(* Logix 5000 project; controller NWGG 1756-L72 rev 35.12; software revision 35.00; part 2 of 19 *)
(* tags used below, declared in another part *)
   T22 : TIMER[100];
   T4 : TIMER[100];

ADD_ON_INSTRUCTION Loadout_K_Valve_Control   (* revision 1.0 *)
VAR_IN_OUT
   K_Valve : udt_Loadout_K_Valve; {required}
   ALM_Clean_Pos_Failed : ALARM_DIGITAL; {required}
   ALM_Treat_Pos_Failed : ALARM_DIGITAL; {required}
   Treat_Position_Input : BOOL; {required}
   Clean_Position_Input : BOOL; {required}
   Clean_Gate_Relay : BOOL; {required}
   Treat_Gate_Relay : BOOL; {required}
END_VAR
VAR
   Clean_Pos_Failed_ACK : BOOL; {access None}
   Treat_Pos_Failedt_ACK : BOOL; {access None}
END_VAR

ROUTINE Logic   (* ladder *)
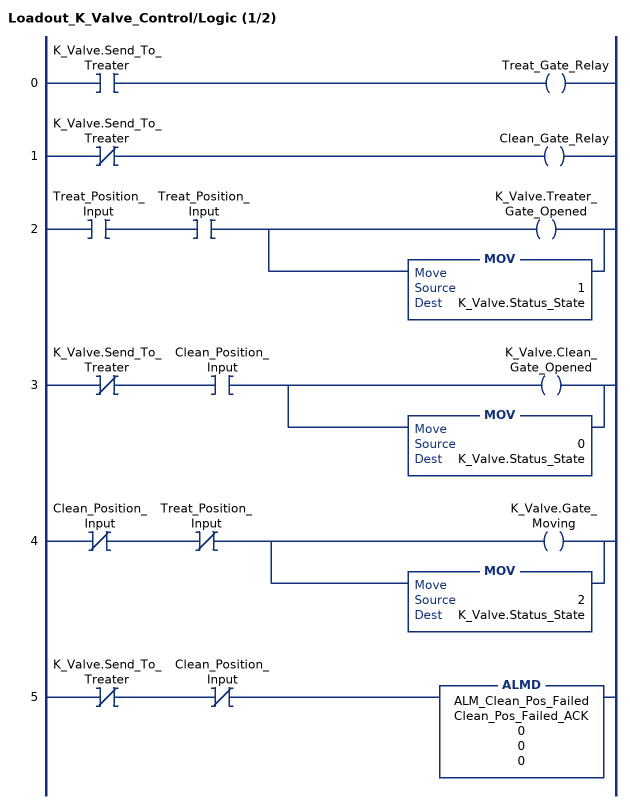
   0: XIC(K_Valve.Send_To_Treater)OTE(Treat_Gate_Relay);
   1: XIO(K_Valve.Send_To_Treater)OTE(Clean_Gate_Relay);
   2: XIC(Treat_Position_Input)XIC(Treat_Position_Input)[OTE(K_Valve.Treater_Gate_Opened) ,MOV(1,K_Valve.Status_State) ];
   3: XIO(K_Valve.Send_To_Treater)XIC(Clean_Position_Input)[OTE(K_Valve.Clean_Gate_Opened) ,MOV(0,K_Valve.Status_State) ];
   4: XIO(Clean_Position_Input)XIO(Treat_Position_Input)[OTE(K_Valve.Gate_Moving) ,MOV(2,K_Valve.Status_State) ];
   5: XIO(K_Valve.Send_To_Treater)XIO(Clean_Position_Input)ALMD(ALM_Clean_Pos_Failed,Clean_Pos_Failed_ACK,0,0,0);
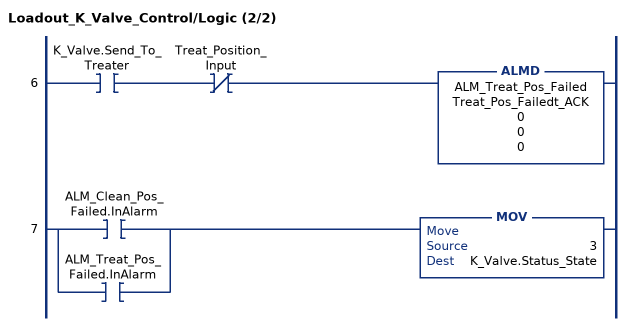
   6: XIC(K_Valve.Send_To_Treater)XIO(Treat_Position_Input)ALMD(ALM_Treat_Pos_Failed,Treat_Pos_Failedt_ACK,0,0,0);
   7: [XIC(ALM_Clean_Pos_Failed.InAlarm) ,XIC(ALM_Treat_Pos_Failed.InAlarm) ]MOV(3,K_Valve.Status_State);
END_ROUTINE
END_ADD_ON_INSTRUCTION

ADD_ON_INSTRUCTION Motor_Control   (* revision 1.0 *)
VAR_IN_OUT
   Motor_Contact : BOOL; {required}
END_VAR
VAR_INPUT
   Spd_20_Pct : BOOL; {required}
   Spd_10_Pct : BOOL; {required}
END_VAR
VAR_OUTPUT
   Running : BOOL; {access Read Only, required}
END_VAR
VAR_IN_OUT
   Motor_Alarm_SPD20 : ALARM_DIGITAL; {required}
   Motor_Alarm_SPD10 : ALARM_DIGITAL; {required}
   Motor_Alarm_Stopped_Over_Amps : ALARM_DIGITAL; {required}
   Motor_Start : udt_Motor_Start; {required}
END_VAR
VAR_INPUT
   Plugged_Sensor : BOOL; {required}
END_VAR
VAR_IN_OUT
   Motor_Alarm_Plugged : ALARM_DIGITAL; {required}
END_VAR
VAR_INPUT
   Motor_Amps : REAL; {required}
END_VAR
VAR_IN_OUT
   Motor_Config : udt_Motor_Config; {required}
   Motor_Starting : BOOL; {required}
   Motor_Alarm_Wont_Start : ALARM_DIGITAL; {required}
END_VAR
VAR_OUTPUT
   In_Alarm : BOOL; {access Read Only}
END_VAR
VAR_IN_OUT
   Treat_Batch_Status : DINT; {required}
   Clean_Batch_Status : DINT; {required}
   Transfer_Batch_Status : DINT; {required}
END_VAR
VAR_OUTPUT
   Motor_Batch_Ready : BOOL; {access Read Only}
END_VAR
VAR_IN_OUT
   Manual_Mode : BOOL; {required}
   InterLocked_Belt : BOOL; {required}
END_VAR
VAR_OUTPUT
   Motor_Batch_Ready_Clean : BOOL; {access Read Only}
   Motor_Batch_Ready_Treat : BOOL; {access Read Only}
   Motor_Batch_Ready_Transfer : BOOL; {access Read Only}
END_VAR
VAR
   TMR_BELT_SPD20 : TIMER := (PRE := 2000); {access None}
   TMR_AMP_INRUSH : TIMER := (PRE := 2000); {access None}
   Alm_Spd20_AK : BOOL; {access None}
   Alm_Spd10_AK : BOOL; {access None}
   Alm_Plugged_AK : BOOL; {access None}
   Alm_OVR_AMP_AK : BOOL; {access None}
   Stop_Motor_Plugged : BOOL; {access None}
   Stop_Motor_SLP20 : BOOL; {access None}
   Stop_Motor : BOOL; {access None}
   Stop_Motor_Ovr_Amp : BOOL; {access None}
   TMR_BELT_SPD10 : TIMER := (PRE := 2000); {access None}
   Alm_Wont_Start_AK : BOOL; {access None}
   Req_Motor_Start : BOOL; {access None}
   tmr_Auto_Stop_Delay : TIMER; {access None}
END_VAR

ROUTINE Logic   (* ladder *)
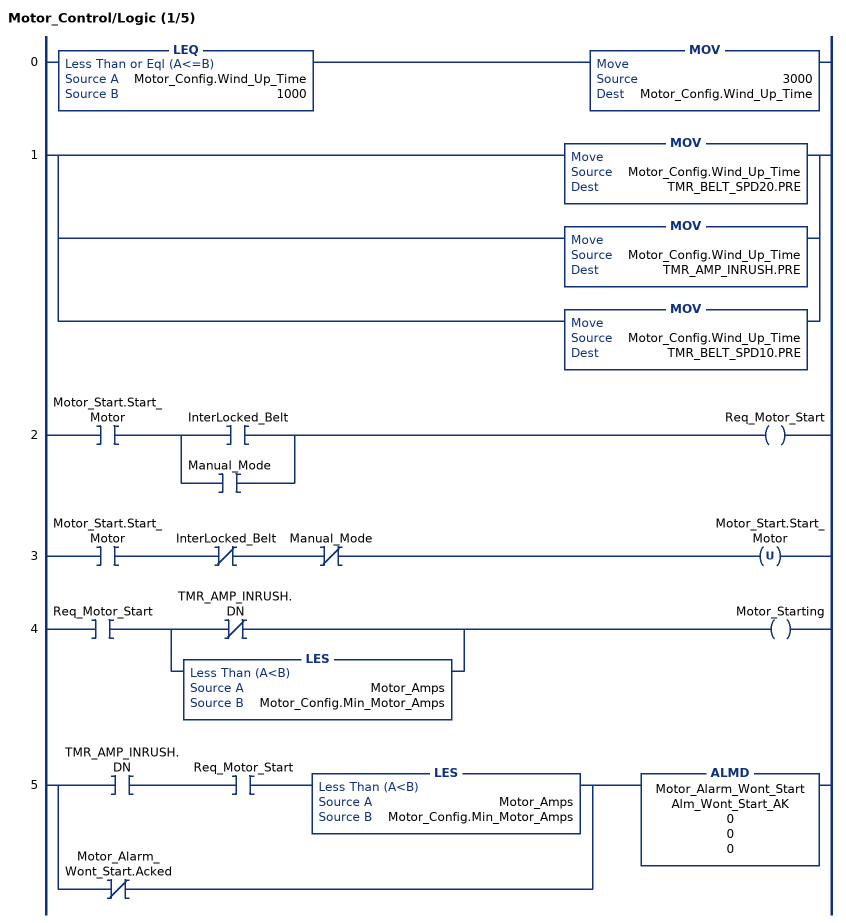
   0: LEQ(Motor_Config.Wind_Up_Time,1000)MOV(3000,Motor_Config.Wind_Up_Time);
   1: [MOV(Motor_Config.Wind_Up_Time,TMR_BELT_SPD20.PRE) ,MOV(Motor_Config.Wind_Up_Time,TMR_AMP_INRUSH.PRE) ,MOV(Motor_Config.Wind_Up_Time,TMR_BELT_SPD10.PRE) ];
   2: XIC(Motor_Start.Start_Motor)[XIC(InterLocked_Belt) ,XIC(Manual_Mode) ]OTE(Req_Motor_Start);
   3: XIC(Motor_Start.Start_Motor)XIO(InterLocked_Belt)XIO(Manual_Mode)OTU(Motor_Start.Start_Motor);
   4: XIC(Req_Motor_Start)[XIO(TMR_AMP_INRUSH.DN) ,LES(Motor_Amps,Motor_Config.Min_Motor_Amps) ]OTE(Motor_Starting);
   5: [XIC(TMR_AMP_INRUSH.DN) XIC(Req_Motor_Start) LES(Motor_Amps,Motor_Config.Min_Motor_Amps) ,XIO(Motor_Alarm_Wont_Start.Acked) ]ALMD(Motor_Alarm_Wont_Start,Alm_Wont_Start_AK,0,0,0);
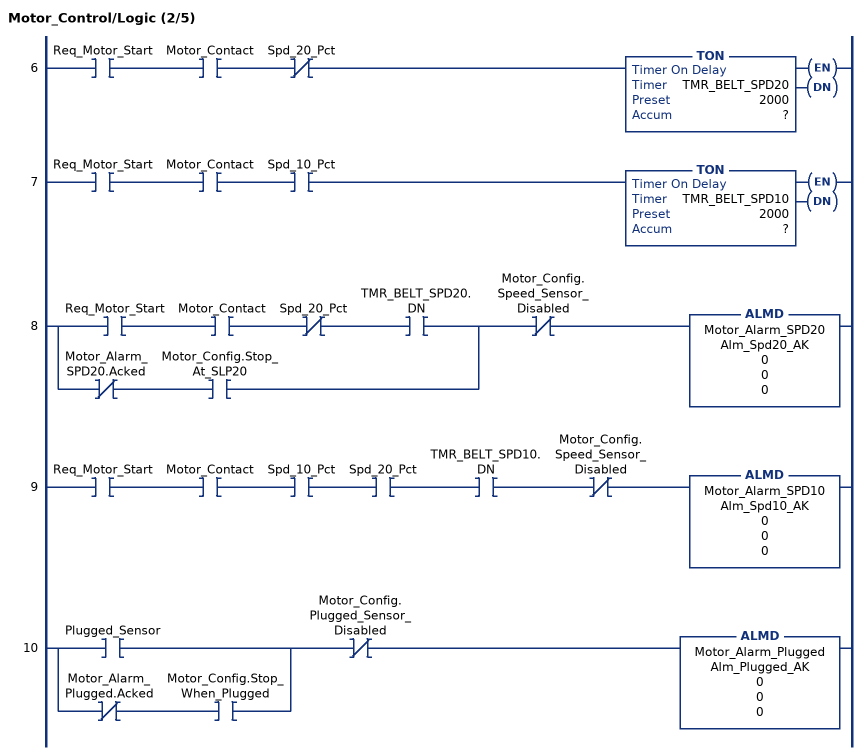
   6: XIC(Req_Motor_Start)XIC(Motor_Contact)XIO(Spd_20_Pct)TON(TMR_BELT_SPD20,?,?);
   7: XIC(Req_Motor_Start)XIC(Motor_Contact)XIC(Spd_10_Pct)TON(TMR_BELT_SPD10,?,?);
   8: [XIC(Req_Motor_Start) XIC(Motor_Contact) XIO(Spd_20_Pct) XIC(TMR_BELT_SPD20.DN) ,XIO(Motor_Alarm_SPD20.Acked) XIC(Motor_Config.Stop_At_SLP20) ]XIO(Motor_Config.Speed_Sensor_Disabled)ALMD(Motor_Alarm_SPD20,Alm_Spd20_AK,0,0,0);
   9: XIC(Req_Motor_Start)XIC(Motor_Contact)XIC(Spd_10_Pct)XIC(Spd_20_Pct)XIC(TMR_BELT_SPD10.DN)XIO(Motor_Config.Speed_Sensor_Disabled)ALMD(Motor_Alarm_SPD10,Alm_Spd10_AK,0,0,0);
   10: [XIC(Plugged_Sensor) ,XIO(Motor_Alarm_Plugged.Acked) XIC(Motor_Config.Stop_When_Plugged) ]XIO(Motor_Config.Plugged_Sensor_Disabled)ALMD(Motor_Alarm_Plugged,Alm_Plugged_AK,0,0,0);
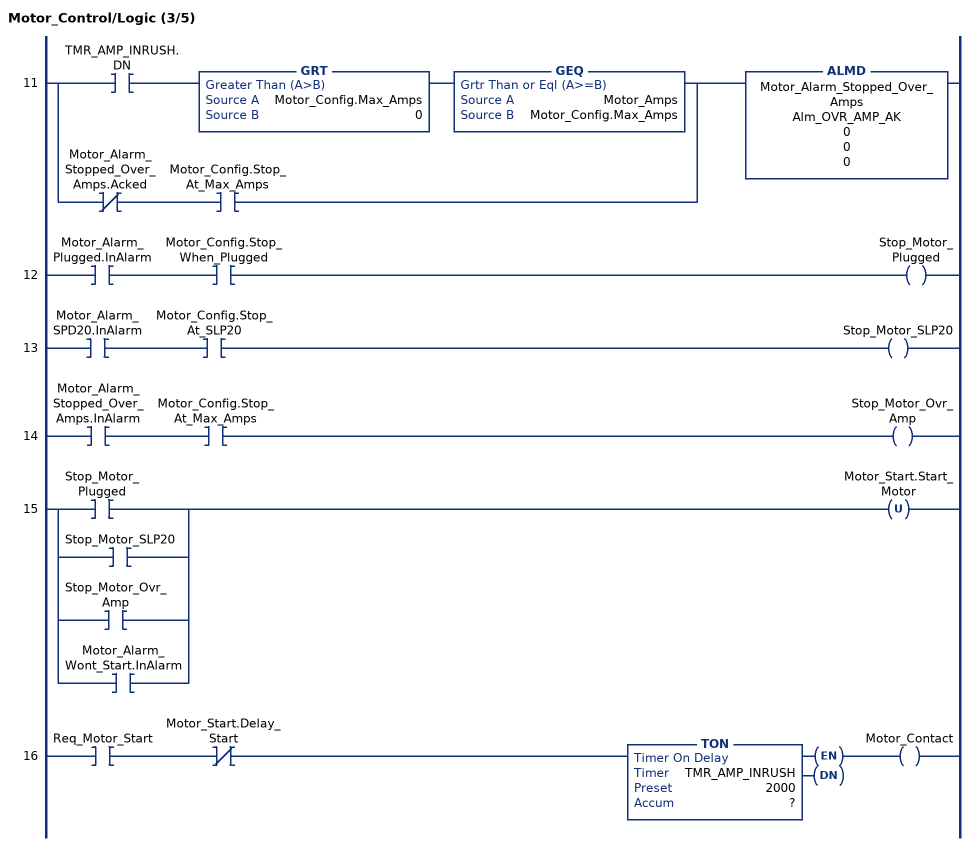
   11: [XIC(TMR_AMP_INRUSH.DN) GRT(Motor_Config.Max_Amps,0) GEQ(Motor_Amps,Motor_Config.Max_Amps) ,XIO(Motor_Alarm_Stopped_Over_Amps.Acked) XIC(Motor_Config.Stop_At_Max_Amps) ]ALMD(Motor_Alarm_Stopped_Over_Amps,Alm_OVR_AMP_AK,0,0,0);
   12: XIC(Motor_Alarm_Plugged.InAlarm)XIC(Motor_Config.Stop_When_Plugged)OTE(Stop_Motor_Plugged);
   13: XIC(Motor_Alarm_SPD20.InAlarm)XIC(Motor_Config.Stop_At_SLP20)OTE(Stop_Motor_SLP20);
   14: XIC(Motor_Alarm_Stopped_Over_Amps.InAlarm)XIC(Motor_Config.Stop_At_Max_Amps)OTE(Stop_Motor_Ovr_Amp);
   15: [XIC(Stop_Motor_Plugged) ,XIC(Stop_Motor_SLP20) ,XIC(Stop_Motor_Ovr_Amp) ,XIC(Motor_Alarm_Wont_Start.InAlarm) ]OTU(Motor_Start.Start_Motor);
   16: XIC(Req_Motor_Start)XIO(Motor_Start.Delay_Start)TON(TMR_AMP_INRUSH,?,?)OTE(Motor_Contact);
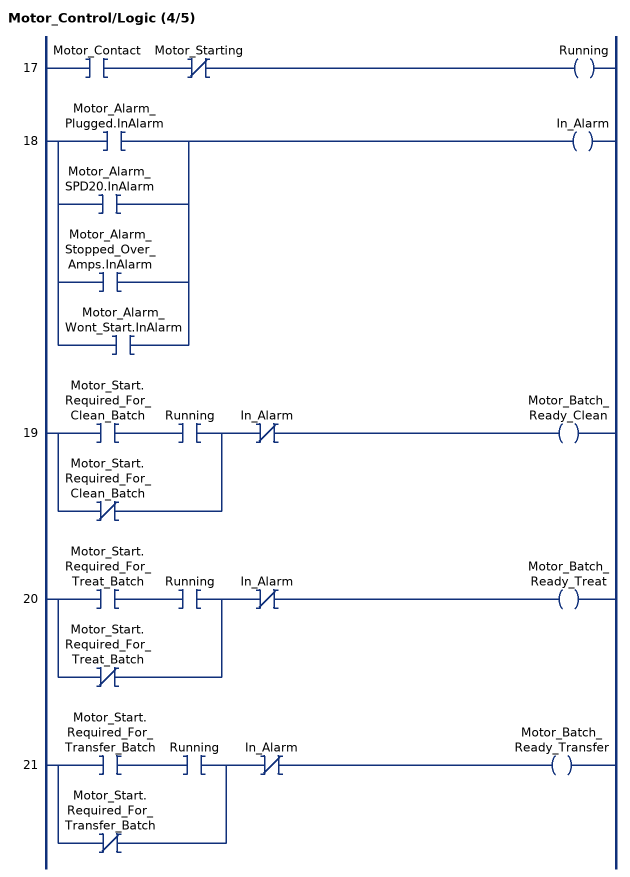
   17: XIC(Motor_Contact)XIO(Motor_Starting)OTE(Running);
   18: [XIC(Motor_Alarm_Plugged.InAlarm) ,XIC(Motor_Alarm_SPD20.InAlarm) ,XIC(Motor_Alarm_Stopped_Over_Amps.InAlarm) ,XIC(Motor_Alarm_Wont_Start.InAlarm) ]OTE(In_Alarm);
   19: [XIC(Motor_Start.Required_For_Clean_Batch) XIC(Running) ,XIO(Motor_Start.Required_For_Clean_Batch) ]XIO(In_Alarm)OTE(Motor_Batch_Ready_Clean);
   20: [XIC(Motor_Start.Required_For_Treat_Batch) XIC(Running) ,XIO(Motor_Start.Required_For_Treat_Batch) ]XIO(In_Alarm)OTE(Motor_Batch_Ready_Treat);
   21: [XIC(Motor_Start.Required_For_Transfer_Batch) XIC(Running) ,XIO(Motor_Start.Required_For_Transfer_Batch) ]XIO(In_Alarm)OTE(Motor_Batch_Ready_Transfer);
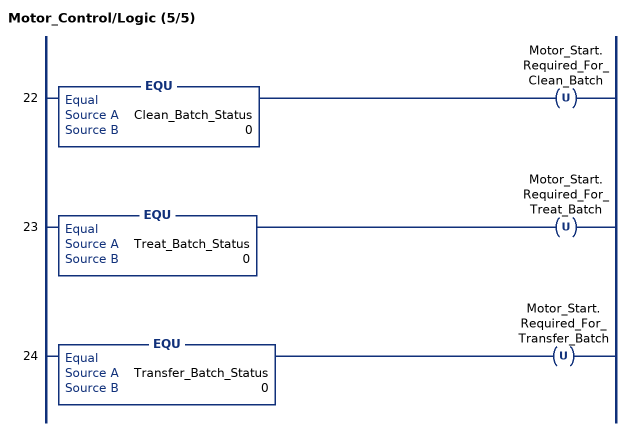
   22: EQU(Clean_Batch_Status,0)OTU(Motor_Start.Required_For_Clean_Batch);
   23: EQU(Treat_Batch_Status,0)OTU(Motor_Start.Required_For_Treat_Batch);
   24: EQU(Transfer_Batch_Status,0)OTU(Motor_Start.Required_For_Transfer_Batch);
END_ROUTINE
END_ADD_ON_INSTRUCTION

ADD_ON_INSTRUCTION SCP   (* revision 1.0, vendor Rockwell Automation *)
VAR_INPUT
   In : ALIAS FOR SCL_01.In; {access None, required}
   InRawMin : REAL; {access None, required}
   InRawMax : REAL; {required}
   InEUMin : REAL; {required}
   InEUMax : REAL; {required}
   Out : DINT; {required}
END_VAR
VAR
   SCL_01 : SCALE; {access None}
   SUB_01 : FBD_MATH; {access None}
   SEL_01 : SELECT; {access None}
   SCL_02 : SCALE; {access None}
   LES_02 : FBD_COMPARE; {access None}
   __l56AFB0E5191E6558 : REAL; {access None}
   __l0BF49CB3D0F7F241 : REAL; {access None}
   __l7339031870541241 : REAL; {access None}
   __l88E0968931849F84 : REAL; {access None}
END_VAR

ROUTINE Logic   (* function block diagram *)
   SHEET 1
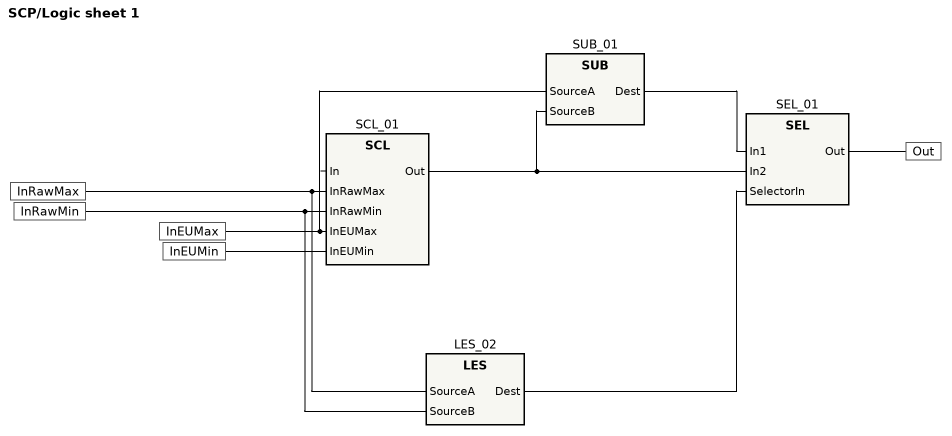
   SCL_01 : SCL(InRawMax := InRawMax, InRawMin := InRawMin, InEUMax := InEUMax, InEUMin := InEUMin);   // unwired pins: In
   LES_02 : LES(SourceA := InRawMax, SourceB := InRawMin);
   SUB_01 : SUB(SourceA := InEUMax, SourceB := SCL_01.Out);
   SEL_01 : SEL(In1 := SUB_01.Dest, In2 := SCL_01.Out, SelectorIn := LES_02.Dest);
   Out := SEL_01.Out;
END_ROUTINE
END_ADD_ON_INSTRUCTION

ADD_ON_INSTRUCTION SCP_Inv   (* revision 1.0, vendor Rockwell Automation *)
VAR_INPUT
   In : ALIAS FOR SCL_01.In; {access None, required}
   InRawMin : REAL; {access None, required}
   InRawMax : REAL; {required}
   InEUMin : REAL; {required}
   InEUMax : REAL; {required}
END_VAR
VAR_OUTPUT
   Out : REAL; {required}
END_VAR
VAR
   SCL_01 : SCALE; {access None}
   SUB_01 : FBD_MATH; {access None}
   SEL_01 : SELECT; {access None}
   SCL_02 : SCALE; {access None}
   LES_02 : FBD_COMPARE; {access None}
   __lC7D96F2B3EA1267C : REAL; {access None}
   __lD4FD1BAAF7FBA06E : REAL; {access None}
   __lFFF49F1C0E6A2B2A : REAL; {access None}
   __lEB05C44F0520614F : REAL; {access None}
END_VAR

ROUTINE Logic   (* function block diagram *)
   SHEET 1
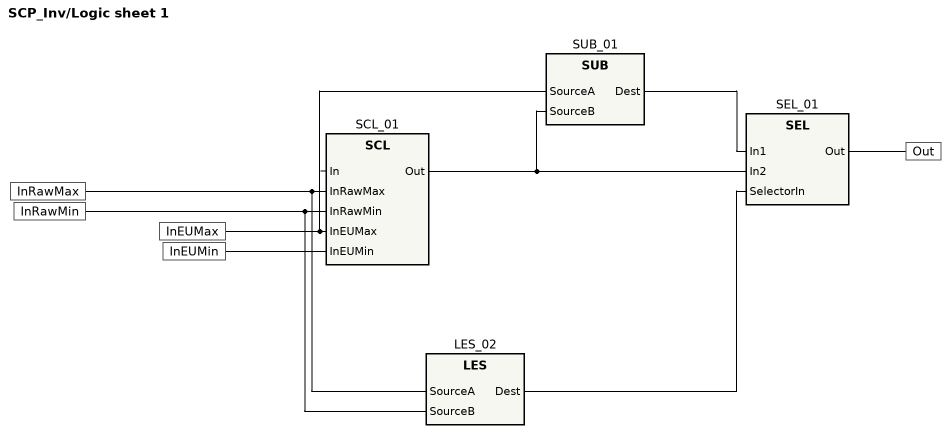
   SCL_01 : SCL(InRawMax := InRawMax, InRawMin := InRawMin, InEUMax := InEUMax, InEUMin := InEUMin);   // unwired pins: In
   LES_02 : LES(SourceA := InRawMax, SourceB := InRawMin);
   SUB_01 : SUB(SourceA := InEUMax, SourceB := SCL_01.Out);
   SEL_01 : SEL(In1 := SUB_01.Dest, In2 := SCL_01.Out, SelectorIn := LES_02.Dest);
   Out := SEL_01.Out;
END_ROUTINE
END_ADD_ON_INSTRUCTION

ADD_ON_INSTRUCTION Truck_Scale_Control   (* revision 1.0 *)
VAR_IN_OUT
   Scale : udt_Truck_Scale; {required}
   Scale_Output : AB:ETHERNET_MODULE_DINT_4Bytes:O:0; {required}
   Scale_Input : AB:ETHERNET_MODULE_DINT_4Bytes:I:0; {required}
END_VAR
VAR
   Rate_Tmr : TIMER := (PRE := 1000, ACC := 713); {access None}
   Accum_Rate_Index1 : COUNTER := (PRE := 11); {access None}
   Old_Accum_Rate : REAL; {access None}
   Rate_Tare : REAL; {access None}
   Lock_Stable_Rate : DINT; {access None}
   Scale_Avg1 : REAL[15]; {access None}
   tmr_Stable : TIMER := (PRE := 2000); {access None}
   tmr_Old_Rate : TIMER := (PRE := 1000); {access None}
   Scale_Avg2 : REAL[15]; {access None}
   Scale_Avg3 : REAL[15]; {access None}
   Avg_Rate1 : REAL; {access None}
   Avg_Rate2 : REAL; {access None}
   Accum_Rate_Index2 : COUNTER := (PRE := 5); {access None}
   Accum_Rate_Index3 : COUNTER := (PRE := 5); {access None}
   Avg_Rate3 : DINT; {access None}
   tmrWeightTest : TIMER; {access None}
END_VAR

ROUTINE Logic   (* ladder *)
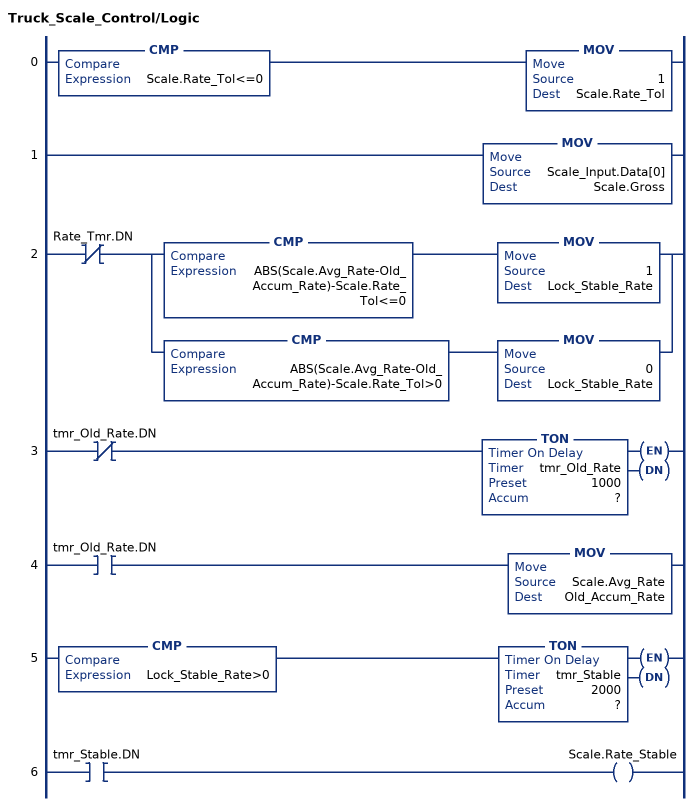
   0: CMP(Scale.Rate_Tol<=0)MOV(1,Scale.Rate_Tol);
   1: MOV(Scale_Input.Data[0],Scale.Gross);
   2: XIO(Rate_Tmr.DN)[CMP(ABS(Scale.Avg_Rate-Old_Accum_Rate)-Scale.Rate_Tol<=0) MOV(1,Lock_Stable_Rate) ,CMP(ABS(Scale.Avg_Rate-Old_Accum_Rate)-Scale.Rate_Tol>0) MOV(0,Lock_Stable_Rate) ];
   3: XIO(tmr_Old_Rate.DN)TON(tmr_Old_Rate,?,?);
   4: XIC(tmr_Old_Rate.DN)MOV(Scale.Avg_Rate,Old_Accum_Rate);
   5: CMP(Lock_Stable_Rate>0)TON(tmr_Stable,?,?);
   6: XIC(tmr_Stable.DN)OTE(Scale.Rate_Stable);
END_ROUTINE
END_ADD_ON_INSTRUCTION

VAR_GLOBAL   (* controller tags *)
   _100AUTO : ALIAS FOR B9[100].4;
   _100HAND : ALIAS FOR B9[100].3;
   _100MB : ALIAS FOR B9[100].2;
   _100STB : ALIAS FOR B9[100].0;
   _100STPB : ALIAS FOR B9[100].1;
   _101_FEED_AUGER_PIT_101_HM : HOUR_METER := (HR_METER_DISPLAY := 21700, MAINTENANCE_ALARM := 1);
   _101AUTO : ALIAS FOR B9[101].4;
   _101HAND : ALIAS FOR B9[101].3;
   _101M : ALIAS FOR O25[9].3;
   _101MB : ALIAS FOR B9[101].2;
   _101STB : ALIAS FOR B9[101].0;
   _101STPB : ALIAS FOR B9[101].1;
   _101Y : ALIAS FOR I25[1].3;
   _102_EXPLORE_TANK_41_RECEIVING_LEG_HM : HOUR_METER := (MOTOR_RUNNING_INPUT_1 := 1, HR_METER_DISPLAY := 13009, MAINTENANCE_ALARM := 1);
   _102AUTO : ALIAS FOR B9[102].4;
   _102HAND : ALIAS FOR B9[102].3;
   _102M : ALIAS FOR O25[8].9;
   _102MB : ALIAS FOR B9[102].2;
   _102STB : ALIAS FOR B9[102].0;
   _102STPB : ALIAS FOR B9[102].1;
   _102Y : ALIAS FOR I25[0].9;
   _103_TANK_42_RECEIVING_LEG_HM : HOUR_METER := (HR_METER_DISPLAY := 4431, NEXT_SCHDL_MAINTENANCE := 2, MAINTENANCE_ALARM := 1);
   _103_TANK_42_RECEIVING_LEG_RUNNING : BOOL;
   _103AUTO : ALIAS FOR B9[103].4;
   _103HAND : ALIAS FOR B9[103].3;
   _103M : ALIAS FOR O25[8].12;
   _103MB : ALIAS FOR B9[103].2;
   _103STB : ALIAS FOR B9[103].0;
   _103STPB : ALIAS FOR B9[103].1;
   _103Y : ALIAS FOR I25[0].12;
   _106_TANK_17_AUGER_HM : HOUR_METER := (HR_METER_DISPLAY := 5679, NEXT_SCHDL_MAINTENANCE := 2, MAINTENANCE_ALARM := 1);
   _106_TANK_17_AUGER_RUNNING : BOOL;
   _106AUTO : ALIAS FOR B9[106].4;
   _106HAND : ALIAS FOR B9[106].3;
   _106M : ALIAS FOR O25[9].5;
   _106MB : ALIAS FOR B9[106].2;
   _106STB : ALIAS FOR B9[106].0;
   _106STPB : ALIAS FOR B9[106].1;
   _106Y : ALIAS FOR I25[1].5;
   _107_SOUTH_BELT_HM : HOUR_METER := (MOTOR_RUNNING_INPUT_1 := 1, HR_METER_DISPLAY := 11100, NEXT_SCHDL_MAINTENANCE := 2, MAINTENANCE_ALARM := 1);
   _107_TANKS_1THRU7_SOUTH_RUNNING : BOOL := 1;
   _107AUTO : ALIAS FOR B9[107].4;
   _107HAND : ALIAS FOR B9[107].3;
   _107M : ALIAS FOR O25[9].12;
   _107MB : ALIAS FOR B9[107].2;
   _107PS : ALIAS FOR I25[4].2;
   _107PSB : ALIAS FOR B9[107].5;
   _107STB : ALIAS FOR B9[107].0;
   _107STPB : ALIAS FOR B9[107].1;
   _107Y : ALIAS FOR I25[1].12;
   _108_CENTER_BELT_HM : HOUR_METER := (MOTOR_RUNNING_INPUT_1 := 1, HR_METER_DISPLAY := 19687, NEXT_SCHDL_MAINTENANCE := 2, MAINTENANCE_ALARM := 1);
   _108_CENTER_BELT_RUNNING : BOOL := 1;
   _108AUTO : ALIAS FOR B9[108].4;
   _108HAND : ALIAS FOR B9[108].3;
   _108M : ALIAS FOR O25[10].15;
   _108MB : ALIAS FOR B9[108].2;
   _108PS : ALIAS FOR I25[4].1;
   _108STB : ALIAS FOR B9[108].0;
   _108STPB : ALIAS FOR B9[108].1;
   _108Y : ALIAS FOR I25[2].15;
   _109_NORTH_BELT_HM : HOUR_METER := (HR_METER_DISPLAY := 77, NEXT_SCHDL_MAINTENANCE := 2, MAINTENANCE_ALARM := 1);
   _109_PS_DLY : ALIAS FOR T11[4];
   _109_RAW_RECEIVING_NORTH_BELT_RUNNING : BOOL;
   _109_SLOW_D : ALIAS FOR T11[5];
   _109_SLW_SP : ALIAS FOR I25[3].14;
   _109_STOP_D : ALIAS FOR T11[6];
   _109_STP_SP : ALIAS FOR I25[3].15;
   _109AUTO : ALIAS FOR B9[109].4;
   _109HAND : ALIAS FOR B9[109].3;
   _109M : ALIAS FOR O25[10].9;
   _109MB : ALIAS FOR B9[109].2;
   _109PS : ALIAS FOR I25[4].0;
   _109STB : ALIAS FOR B9[109].0;
   _109STPB : ALIAS FOR B9[109].1;
   _109Y : ALIAS FOR I25[2].9;
   _10AUTO : ALIAS FOR B9[10].4;
   _10HAND : ALIAS FOR B9[10].3;
   _10MB : ALIAS FOR B9[10].2;
   _10STB : ALIAS FOR B9[10].0;
   _10STPB : ALIAS FOR B9[10].1;
   _10Y : ALIAS FOR I25[0].11;
   _110_TANK_16_AUGER_HM : HOUR_METER := (HR_METER_DISPLAY := 3779, NEXT_SCHDL_MAINTENANCE := 2, MAINTENANCE_ALARM := 1);
   _110_TANK_16_AUGER_RUNNING : BOOL;
   _110AUTO : ALIAS FOR B9[110].4;
   _110HAND : ALIAS FOR B9[110].3;
   _110M : ALIAS FOR O25[8].15;
   _110MB : ALIAS FOR B9[110].2;
   _110STB : ALIAS FOR B9[110].0;
   _110STPB : ALIAS FOR B9[110].1;
   _110Y : ALIAS FOR I25[0].15;
   _111_TANK_17_AUGER_HM : HOUR_METER := (HR_METER_DISPLAY := 1055, MAINTENANCE_ALARM := 1);
   _111AUTO : ALIAS FOR B9[111].4;
   _111HAND : ALIAS FOR B9[111].3;
   _111M : ALIAS FOR O25[9].0;
   _111MB : ALIAS FOR B9[111].2;
   _111STB : ALIAS FOR B9[111].0;
   _111STPB : ALIAS FOR B9[111].1;
   _111Y : ALIAS FOR I25[1].0;
   _113_GATE_B : ALIAS FOR I25[4].12;
   _113_GATE_B1 : ALIAS FOR I25[4].13;
   _113_HIGHROLLER_TANKS_11TO15_HM : HOUR_METER := (HR_METER_DISPLAY := 1063, NEXT_SCHDL_MAINTENANCE := 2, MAINTENANCE_ALARM := 1);
   _113_HIGHROLLER_TANKS_11TO15_RUNNING : BOOL;
   _113_TO_BC1 : ALIAS FOR O25[11].9;
   _113_TO_BC9 : ALIAS FOR O25[11].8;
   _113AUTO : ALIAS FOR B9[113].4;
   _113HAND : ALIAS FOR B9[113].3;
   _113M : ALIAS FOR O25[10].5;
   _113MB : ALIAS FOR B9[113].2;
   _113STB : ALIAS FOR B9[113].0;
   _113STPB : ALIAS FOR B9[113].1;
   _113Y : ALIAS FOR I25[2].5;
   _114_TANKS_1THRU7_NORTH_HM : HOUR_METER := (HR_METER_DISPLAY := 9528, MAINTENANCE_ALARM := 1);
   _114_TANKS_1THRU7_NORTH_RUNNING : BOOL;
   _115_M : ALIAS FOR O25[22].0;
   _115AUTO : ALIAS FOR B9[115].4;
   _115HAND : ALIAS FOR B9[115].3;
   _115MB : ALIAS FOR B9[115].2;
   _115STB : ALIAS FOR B9[115].0;
   _115STPB : ALIAS FOR B9[115].1;
   _116_DRAG_16_HM : HOUR_METER := (HR_METER_DISPLAY := 3781, MAINTENANCE_ALARM := 1);
   _116AUTO : ALIAS FOR B9[116].4;
   _116HAND : ALIAS FOR B9[116].3;
   _116M : ALIAS FOR O25[10].10;
   _116MB : ALIAS FOR B9[116].2;
   _116STB : ALIAS FOR B9[116].0;
   _116STPB : ALIAS FOR B9[116].1;
   _116Y : ALIAS FOR I25[2].10;
   _117_DRAG_17_HM : HOUR_METER := (HR_METER_DISPLAY := 5681, MAINTENANCE_ALARM := 1);
   _117AUTO : ALIAS FOR B9[117].4;
   _117HAND : ALIAS FOR B9[117].3;
   _117M : ALIAS FOR O25[10].8;
   _117MB : ALIAS FOR B9[117].2;
   _117STB : ALIAS FOR B9[117].0;
   _117STPB : ALIAS FOR B9[117].1;
   _117Y : ALIAS FOR I25[2].8;
   _11_BINDICA : ALIAS FOR B15[11].0;
   _11_BINDICA1 : ALIAS FOR B15[11].1;
   _11_GATE_PO : ALIAS FOR I16[0];
   _11_GATE_PO1 : ALIAS FOR N14[11];
   _11_GATE_PO_STOR : REAL := 86.33458;
   _11_PS : ALIAS FOR I25[4].14;
   _11_PS_DLY : ALIAS FOR T11[2];
   _11_SLOW_SP : ALIAS FOR I25[4].3;
   _11_STOP_SP : ALIAS FOR I25[4].6;
   _11_TANK_41_42_HIGHROLLER_HM : HOUR_METER := (HR_METER_DISPLAY := 6844, NEXT_SCHDL_MAINTENANCE := 2, MAINTENANCE_ALARM := 1);
   _11_TANK_41_42_HIGHROLLER_RUNNING : BOOL;
   _11_VALVE_R : ALIAS FOR I25[4].4;
   _11_VALVE_S : ALIAS FOR I25[4].5;
   _11AUTO : ALIAS FOR B9[11].4;
   _11HAND : ALIAS FOR B9[11].3;
   _11M : ALIAS FOR O25[9].2;
   _11MB : ALIAS FOR B9[11].2;
   _11STB : ALIAS FOR B9[11].0;
   _11STPB : ALIAS FOR B9[11].1;
   _11Y : ALIAS FOR I25[1].2;
   _122_RECIEVING_LEG_HM : HOUR_METER := (MOTOR_RUNNING_INPUT_1 := 1, HR_METER_DISPLAY := 24537, MAINTENANCE_ALARM := 1);
   _122AUTO : ALIAS FOR B9[122].4;
   _122HAND : ALIAS FOR B9[122].3;
   _122M : ALIAS FOR O25[9].1;
   _122MB : ALIAS FOR B9[122].2;
   _122STB : ALIAS FOR B9[122].0;
   _122STPB : ALIAS FOR B9[122].1;
   _122Y : ALIAS FOR I25[1].1;
   _123_CLEAN_LEG_HM : HOUR_METER := (MOTOR_RUNNING_INPUT_1 := 1, HR_METER_DISPLAY := 26622, NEXT_SCHDL_MAINTENANCE := 2, MAINTENANCE_ALARM := 1);
   _123_CLEAN_LEG_RUNNING : BOOL := 1;
   _123_COMPUW : ALIAS FOR I18[7];
   _123_COMPUW1 : ALIAS FOR N7[20];
   _123AUTO : ALIAS FOR B9[123].4;
   _123HAND : ALIAS FOR B9[123].3;
   _123M : ALIAS FOR O25[10].6;
   _123MB : ALIAS FOR B9[123].2;
   _123STB : ALIAS FOR B9[123].0;
   _123STPB : ALIAS FOR B9[123].1;
   _123Y : ALIAS FOR I25[2].6;
   _124AUTO : ALIAS FOR B9[124].4;
   _124HAND : ALIAS FOR B9[124].3;
   _124M : ALIAS FOR O25[9].13;
   _124MB : ALIAS FOR B9[124].2;
   _124STB : ALIAS FOR B9[124].0;
   _124STPB : ALIAS FOR B9[124].1;
   _125_COLOR_SORTER_LEG_HM : HOUR_METER := (MOTOR_RUNNING_INPUT_1 := 1, HR_METER_DISPLAY := 26513, NEXT_SCHDL_MAINTENANCE := 2, MAINTENANCE_ALARM := 1);
   _126_ASPERATOR : HOUR_METER := (MOTOR_RUNNING_INPUT_1 := 1, HR_METER_DISPLAY := 25758, NEXT_SCHDL_MAINTENANCE := 2, MAINTENANCE_ALARM := 1);
   _128_SCREENINGS_DRAG_HM : HOUR_METER := (MOTOR_RUNNING_INPUT_1 := 1, HR_METER_DISPLAY := 26532, NEXT_SCHDL_MAINTENANCE := 2, MAINTENANCE_ALARM := 1);
   _12_BINDICA : ALIAS FOR B15[12].0;
   _12_BINDICA1 : ALIAS FOR B15[12].1;
   _12_GATE_PO : ALIAS FOR I16[1];
   _12_GATE_PO1 : ALIAS FOR N14[12];
   _12_GATE_PO_STOR : REAL := 94.72872;
   _13_BINDICA : ALIAS FOR B15[13].0;
   _13_BINDICA1 : ALIAS FOR B15[13].1;
   _13_GATE_PO : ALIAS FOR I16[2];
   _13_GATE_PO1 : ALIAS FOR N14[13];
   _13_GATE_PO_STOR : REAL := 79.42468;
   _14_BINDICA : ALIAS FOR B15[14].0;
   _14_BINDICA1 : ALIAS FOR B15[14].1;
   _14_GATE_PO : ALIAS FOR I16[3];
   _14_GATE_PO1 : ALIAS FOR N14[14];
   _14_GATE_PO_STOR : REAL := 93.90426;
   _15_BINDICA : ALIAS FOR B15[15].0;
   _15_BINDICA1 : ALIAS FOR B15[15].1;
   _15_GATE_PO : ALIAS FOR I16[4];
   _15_GATE_PO1 : ALIAS FOR N14[15];
   _15_GATE_PO_STOR : REAL := 92.96653;
   _16_BINDICA : ALIAS FOR B15[16].0;
   _16_BINDICA1 : ALIAS FOR B15[16].1;
   _16_GATE_PO : ALIAS FOR I16[5];
   _16_GATE_PO1 : ALIAS FOR N14[16];
   _16_GATE_PO_STOR : REAL := 30.742159;
   _17_BINDICA : ALIAS FOR B15[17].0;
   _17_BINDICA1 : ALIAS FOR B15[17].1;
   _17_GATE_PO : ALIAS FOR I16[6];
   _17_GATE_PO1 : ALIAS FOR N14[17];
   _17_GATE_PO_STOR : REAL := 78.57861;
   _1_CLEAN_SEED_UPPER_BELT_HM : HOUR_METER := (MOTOR_RUNNING_INPUT_1 := 1, HR_METER_DISPLAY := 13589, NEXT_SCHDL_MAINTENANCE := 2, MAINTENANCE_ALARM := 1);
   _1_CLEAN_SEED_UPPER_BELT_RUNNING : BOOL := 1;
   _1AUTO : ALIAS FOR B9[1].4;
   _1HAND : ALIAS FOR B9[1].3;
   _1M : ALIAS FOR O25[9].8;
   _1MB : ALIAS FOR B9[1].2;
   _1STB : ALIAS FOR B9[1].0;
   _1STPB : ALIAS FOR B9[1].1;
   _1Y : ALIAS FOR I25[1].8;
   _21_BINDICA : ALIAS FOR B15[21].0;
   _21_BINDICA1 : ALIAS FOR B15[21].1;
   _21_GATE_PO : ALIAS FOR I16[7];
   _21_GATE_PO1 : ALIAS FOR N14[21];
   _21_GATE_PO_STOR : REAL := 87.275024;
   _22_BINDICA : ALIAS FOR B15[22].0;
   _22_BINDICA1 : ALIAS FOR B15[22].1;
   _22_GATE_PO : ALIAS FOR I17[0];
   _22_GATE_PO1 : ALIAS FOR N14[22];
   _22_GATE_PO_STOR : REAL := 83.08857;
   _22AUTO : ALIAS FOR B9[22].4;
   _22HAND : ALIAS FOR B9[22].3;
   _22MB : ALIAS FOR B9[22].2;
   _22STB : ALIAS FOR B9[22].0;
   _22STPB : ALIAS FOR B9[22].1;
   _23_BINDICA : ALIAS FOR B15[23].0;
   _23_BINDICA1 : ALIAS FOR B15[23].1;
   _23_GATE_PO : ALIAS FOR I17[1];
   _23_GATE_PO1 : ALIAS FOR N14[23];
   _23_GATE_PO_STOR : REAL := 96.74677;
   _24_16_0 : ALIAS FOR N250[0];
   _24_16_1 : ALIAS FOR N250[1];
   _24_16_2 : ALIAS FOR N250[2];
   _24_16_3 : ALIAS FOR N250[3];
   _24_16_4 : ALIAS FOR N250[4];
   _24_16_5 : ALIAS FOR N250[5];
   _24_16_6 : ALIAS FOR N250[6];
   _24_16_7 : ALIAS FOR N250[7];
   _24_16_BLK : ALIAS FOR T4[58];
   _24_17_0 : ALIAS FOR N240[0];
   _24_17_1 : ALIAS FOR N240[1];
   _24_17_2 : ALIAS FOR N240[2];
   _24_17_3 : ALIAS FOR N240[3];
   _24_17_4 : ALIAS FOR N240[4];
   _24_17_5 : ALIAS FOR N240[5];
   _24_17_6 : ALIAS FOR N240[6];
   _24_17_7 : ALIAS FOR N240[7];
   _24_17_BLK : ALIAS FOR T4[57];
   _24_18_0_AN : ALIAS FOR N230[10];
   _24_18_1_AN : ALIAS FOR N230[11];
   _24_18_2_AN : ALIAS FOR N230[12];
   _24_18_3_AN : ALIAS FOR N230[13];
   _24_18_BLK : ALIAS FOR T4[40];
   _24_18_MULT : ALIAS FOR N230[14];
   _24_19_0 : ALIAS FOR N220[10];
   _24_19_1 : ALIAS FOR N220[11];
   _24_19_2 : ALIAS FOR N220[12];
   _24_19_3 : ALIAS FOR N220[13];
   _24_19_BLK : ALIAS FOR T4[39];
   _24_20_0 : ALIAS FOR N210[10];
   _24_20_1 : ALIAS FOR N210[11];
   _24_20_2 : ALIAS FOR N210[12];
   _24_20_3 : ALIAS FOR N210[13];
   _24_20_BLK : ALIAS FOR T4[38];
   _24_BINDICA : ALIAS FOR B15[24].0;
   _24_BINDICA1 : ALIAS FOR B15[24].1;
   _24_GATE_PO : ALIAS FOR I17[2];
   _24_GATE_PO1 : ALIAS FOR N14[24];
   _24_GATE_PO_STOR : REAL := 90.36168;
   _25_16_0 : ALIAS FOR N200[10];
   _25_16_1 : ALIAS FOR N200[11];
   _25_16_2 : ALIAS FOR N200[12];
   _25_16_3 : ALIAS FOR N200[13];
   _25_16_BLK : ALIAS FOR T4[37];
   _25_17_0 : ALIAS FOR N190[0];
   _25_17_1 : ALIAS FOR N190[1];
   _25_17_2 : ALIAS FOR N190[2];
   _25_17_3 : ALIAS FOR N190[3];
   _25_17_BLK : ALIAS FOR T4[36];
   _25_18_TMR : ALIAS FOR T4[35];
   _25_BINDICA : ALIAS FOR B15[25].0;
   _25_BINDICA1 : ALIAS FOR B15[25].1;
   _25_GATE_PO : ALIAS FOR I17[3];
   _25_GATE_PO1 : ALIAS FOR N14[25];
   _25_GATE_PO_STOR : REAL := 103.03115;
   _26_BINDICA : ALIAS FOR B15[26].0;
   _26_BINDICA1 : ALIAS FOR B15[26].1;
   _26_GATE_PO : ALIAS FOR I17[4];
   _26_GATE_PO1 : ALIAS FOR N14[26];
   _26_GATE_PO_STOR : REAL := 98.9571;
   _27_BINDICA : ALIAS FOR B15[27].0;
   _27_BINDICA1 : ALIAS FOR B15[27].1;
   _27_GATE_PO : ALIAS FOR I17[5];
   _27_GATE_PO1 : ALIAS FOR N14[27];
   _28_BINDICA : ALIAS FOR B15[28].0;
   _28_BINDICA1 : ALIAS FOR B15[28].1;
   _28_GATE_PO : ALIAS FOR I17[6];
   _28_GATE_PO1 : ALIAS FOR N14[28];
   _29_BINDICA : ALIAS FOR B15[29].0;
   _29_BINDICA1 : ALIAS FOR B15[29].1;
   _29_GATE_PO : ALIAS FOR I17[7];
   _29_GATE_PO1 : ALIAS FOR N14[29];
   _2AUTO : ALIAS FOR B9[2].4;
   _2HAND : ALIAS FOR B9[2].3;
   _2M : ALIAS FOR O25[9].15;
   _2MB : ALIAS FOR B9[2].2;
   _2STB : ALIAS FOR B9[2].0;
   _2STPB : ALIAS FOR B9[2].1;
   _2Y : ALIAS FOR I25[1].15;
   _35_JUMP_LEG_HM : HOUR_METER := (MOTOR_RUNNING_INPUT_1 := 1, HR_METER_DISPLAY := 26389, NEXT_SCHDL_MAINTENANCE := 2, MAINTENANCE_ALARM := 1);
   _35_JUMP_LEG_RUNNING : BOOL := 1;
   _35AUTO : ALIAS FOR B9[35].4;
   _35HAND : ALIAS FOR B9[35].3;
   _35M : ALIAS FOR O25[10].13;
   _35MB : ALIAS FOR B9[35].2;
   _35STB : ALIAS FOR B9[35].0;
   _35STPB : ALIAS FOR B9[35].1;
   _35Y : ALIAS FOR I25[2].13;
   _36_FREQ_IN : ALIAS FOR N7[1];
   _36_FREQ_OU : ALIAS FOR N7[3];
   _36_SET_SPD : ALIAS FOR N7[2];
   _36_TANK_41_AUGER_HM : HOUR_METER := (HR_METER_DISPLAY := 2995, MAINTENANCE_ALARM := 1);
   _36_VFD_TO : ALIAS FOR N180[0];
   _36M : ALIAS FOR O25[8].0;
   _36MAI : ALIAS FOR O25[25].0;
   _36RAUTO : ALIAS FOR B9[36].4;
   _36RHAND : ALIAS FOR B9[36].3;
   _36RMB : ALIAS FOR B9[36].2;
   _36RSTB : ALIAS FOR B9[36].0;
   _36RSTPB : ALIAS FOR B9[36].1;
   _36RY : ALIAS FOR I25[16].0;
   _36Y : ALIAS FOR I25[0].0;
   _3_LOWER_TANK_CONVAYOR_24TO26_HM : HOUR_METER := (HR_METER_DISPLAY := 1012, NEXT_SCHDL_MAINTENANCE := 2, MAINTENANCE_ALARM := 1);
   _3_LOWER_TANK_CONVAYOR_24TO26_RUNNING : BOOL;
   _3_LS_TO_5 : ALIAS FOR I25[4].8;
   _3_LS_TO_6 : ALIAS FOR I25[4].9;
   _3_TO_BC5_S : ALIAS FOR O25[11].12;
   _3_TO_BC6_S : ALIAS FOR O25[11].13;
   _3AUTO : ALIAS FOR B9[3].4;
   _3HAND : ALIAS FOR B9[3].3;
   _3M : ALIAS FOR O25[10].0;
   _3MB : ALIAS FOR B9[3].2;
   _3STB : ALIAS FOR B9[3].0;
   _3STPB : ALIAS FOR B9[3].1;
   _3Y : ALIAS FOR I25[2].0;
   _41_GATE_PO : ALIAS FOR I18[0];
   _41_GATE_PO1 : ALIAS FOR N14[41];
   _42_GATE_PO : ALIAS FOR I18[1];
   _42_GATE_PO1 : ALIAS FOR N14[42];
   _42_LOWER_SCREENINGS_DRAG_HM : HOUR_METER := (MOTOR_RUNNING_INPUT_1 := 1, HR_METER_DISPLAY := 27637, MAINTENANCE_ALARM := 1);
   _42AUTO : ALIAS FOR B9[42].4;
   _42HAND : ALIAS FOR B9[42].3;
   _42M : ALIAS FOR O25[11].1;
   _42MB : ALIAS FOR B9[42].2;
   _42STB : ALIAS FOR B9[42].0;
   _42STPB : ALIAS FOR B9[42].1;
   _42Y : ALIAS FOR I25[3].1;
   _43_ACC_WEI : ALIAS FOR C5[1].ACC;
   _43_BINDICA : ALIAS FOR B9[43].5;
   _43_RESET_C : ALIAS FOR B9[43].6;
   _43_SCREEN : ALIAS FOR C5[1];
   _43_SCREENI : ALIAS FOR I7.14;
   _43_SCREENINGS_LEG_HM : HOUR_METER := (MOTOR_RUNNING_INPUT_1 := 1, HR_METER_DISPLAY := 27656, NEXT_SCHDL_MAINTENANCE := 2, MAINTENANCE_ALARM := 1);
   _43_SCREENINGS_LEG_RUNNING : BOOL := 1;
   _43_WEIGHT : ALIAS FOR N7[0];
   _43AUTO : ALIAS FOR B9[43].4;
   _43HAND : ALIAS FOR B9[43].3;
   _43M : ALIAS FOR O25[10].14;
   _43MB : ALIAS FOR B9[43].2;
   _43STB : ALIAS FOR B9[43].0;
   _43STPB : ALIAS FOR B9[43].1;
   _43Y : ALIAS FOR I25[2].14;
   _45_AIR_SEQ : ALIAS FOR T4[34];
   _45_AIR_SEQ1 : ALIAS FOR T4[34].PRE;
   _45_AIR_SEQ2 : ALIAS FOR T4[34].ACC;
   _45_SEQ_AIR : ALIAS FOR O12.15;
   _45AUTO : ALIAS FOR B9[45].4;
   _45HAND : ALIAS FOR B9[45].3;
   _45M : ALIAS FOR O25[8].7;
   _45MB : ALIAS FOR B9[45].2;
   _45STB : ALIAS FOR B9[45].0;
   _45STPB : ALIAS FOR B9[45].1;
   _45Y : ALIAS FOR I25[0].7;
   _46AUTO : ALIAS FOR B9[46].4;
   _46HAND : ALIAS FOR B9[46].3;
   _46M : ALIAS FOR O25[8].8;
   _46MB : ALIAS FOR B9[46].2;
   _46STB : ALIAS FOR B9[46].0;
   _46STPB : ALIAS FOR B9[46].1;
   _46Y : ALIAS FOR I25[0].8;
   _47AUTO : ALIAS FOR B9[47].4;
   _47HAND : ALIAS FOR B9[47].3;
   _47M : ALIAS FOR O25[9].10;
   _47MB : ALIAS FOR B9[47].2;
   _47STB : ALIAS FOR B9[47].0;
   _47STPB : ALIAS FOR B9[47].1;
   _47Y : ALIAS FOR I25[1].10;
   _48_CIMBRIA_HM : HOUR_METER := (MOTOR_RUNNING_INPUT_1 := 1, HR_METER_DISPLAY := 24757, MAINTENANCE_ALARM := 1);
   _48_FREQ_IN : ALIAS FOR N7[10];
   _48_FREQ_OU : ALIAS FOR N7[12];
   _48_SET_SPD : ALIAS FOR N7[11];
   _48_VFD_TO : ALIAS FOR N180[2];
   _48AUTO : ALIAS FOR B9[48].4;
   _48HAND : ALIAS FOR B9[48].3;
   _48M : ALIAS FOR O25[8].3;
   _48MAI : ALIAS FOR O25[25].2;
   _48MB : ALIAS FOR B9[48].2;
   _48STB : ALIAS FOR B9[48].0;
   _48STPB : ALIAS FOR B9[48].1;
   _48Y : ALIAS FOR I25[0].3;
   _49AUTO : ALIAS FOR B9[49].4;
   _49HAND : ALIAS FOR B9[49].3;
   _49M : ALIAS FOR O25[9].9;
   _49MB : ALIAS FOR B9[49].2;
   _49STB : ALIAS FOR B9[49].0;
   _49STPB : ALIAS FOR B9[49].1;
   _49Y : ALIAS FOR I25[1].9;
   _4_LOWER_TANK_CONVAYOR_21TO23_HM : HOUR_METER := (HR_METER_DISPLAY := 1470, NEXT_SCHDL_MAINTENANCE := 2, MAINTENANCE_ALARM := 1);
   _4_LOWER_TANK_CONVAYOR_21TO23_RUNNING : BOOL;
   _4_LS_TO_5 : ALIAS FOR I25[4].10;
   _4_LS_TO_6 : ALIAS FOR I25[4].11;
   _4_TO_BC5_S : ALIAS FOR O25[11].10;
   _4_TO_BC6_S : ALIAS FOR O25[11].11;
   _4AUTO : ALIAS FOR B9[4].4;
   _4HAND : ALIAS FOR B9[4].3;
   _4M : ALIAS FOR O25[10].1;
   _4MB : ALIAS FOR B9[4].2;
   _4STB : ALIAS FOR B9[4].0;
   _4STPB : ALIAS FOR B9[4].1;
   _4Y : ALIAS FOR I25[2].1;
   _50AUTO : ALIAS FOR B9[50].4;
   _50HAND : ALIAS FOR B9[50].3;
   _50M : ALIAS FOR O25[8].14;
   _50MB : ALIAS FOR B9[50].2;
   _50STB : ALIAS FOR B9[50].0;
   _50STPB : ALIAS FOR B9[50].1;
   _50Y : ALIAS FOR I25[0].14;
   _51_FREQ_IN : ALIAS FOR N7[13];
   _51_FREQ_OU : ALIAS FOR N7[15];
   _51_INDENT_HM : HOUR_METER := (MOTOR_RUNNING_INPUT_1 := 1, HR_METER_DISPLAY := 26515, MAINTENANCE_ALARM := 1);
   _51_SET_SPD : ALIAS FOR N7[14];
   _51_VFD_TO : ALIAS FOR N180[3];
   _51AUTO : ALIAS FOR B9[51].4;
   _51HAND : ALIAS FOR B9[51].3;
   _51M : ALIAS FOR O25[8].4;
   _51MAI : ALIAS FOR O25[25].3;
   _51MB : ALIAS FOR B9[51].2;
   _51STB : ALIAS FOR B9[51].0;
   _51STPB : ALIAS FOR B9[51].1;
   _51Y : ALIAS FOR I25[0].4;
   _52_FREQ_IN : ALIAS FOR N7[16];
   _52_FREQ_OU : ALIAS FOR N7[18];
   _52_SET_SPD : ALIAS FOR N7[17];
   _52AUTO : ALIAS FOR B9[52].4;
   _52HAND : ALIAS FOR B9[52].3;
   _52M : ALIAS FOR O25[8].6;
   _52MAI : ALIAS FOR O25[25].4;
   _52MB : ALIAS FOR B9[52].2;
   _52STB : ALIAS FOR B9[52].0;
   _52STPB : ALIAS FOR B9[52].1;
   _52Y : ALIAS FOR I25[0].6;
   _53_FREQ_IN : ALIAS FOR N7[7];
   _53_FREQ_OU : ALIAS FOR N7[9];
   _53_SET_SPD : ALIAS FOR N7[8];
   _53_VFD_TO : ALIAS FOR N180[1];
   _53AUTO : ALIAS FOR B9[53].4;
   _53HAND : ALIAS FOR B9[53].3;
   _53M : ALIAS FOR O25[8].2;
   _53MAI : ALIAS FOR O25[25].1;
   _53MB : ALIAS FOR B9[53].2;
   _53STB : ALIAS FOR B9[53].0;
   _53STPB : ALIAS FOR B9[53].1;
   _53Y : ALIAS FOR I25[0].2;
   _54AUTO : ALIAS FOR B9[54].4;
   _54HAND : ALIAS FOR B9[54].3;
   _54M : ALIAS FOR O25[11].3;
   _54MB : ALIAS FOR B9[54].2;
   _54STB : ALIAS FOR B9[54].0;
   _54STPB : ALIAS FOR B9[54].1;
   _54Y : ALIAS FOR I25[3].3;
   _55_FREQ_IN : ALIAS FOR N7[4];
   _55_FREQ_OU : ALIAS FOR N7[6];
   _55_SET_SPD : ALIAS FOR N7[5];
   _55AUTO : ALIAS FOR B9[55].4;
   _55HAND : ALIAS FOR B9[55].3;
   _55M : ALIAS FOR O25[8].1;
   _55MB : ALIAS FOR B9[55].2;
   _55STB : ALIAS FOR B9[55].0;
   _55STPB : ALIAS FOR B9[55].1;
   _55Y : ALIAS FOR I25[0].1;
   _56AUTO : ALIAS FOR B9[56].4;
   _56HAND : ALIAS FOR B9[56].3;
   _56M : ALIAS FOR O25[11].2;
   _56MB : ALIAS FOR B9[56].2;
   _56STB : ALIAS FOR B9[56].0;
   _56STPB : ALIAS FOR B9[56].1;
   _56Y : ALIAS FOR I25[3].2;
   _57AUTO : ALIAS FOR B9[57].4;
   _57HAND : ALIAS FOR B9[57].3;
   _57M : ALIAS FOR O25[9].6;
   _57MB : ALIAS FOR B9[57].2;
   _57STB : ALIAS FOR B9[57].0;
   _57STPB : ALIAS FOR B9[57].1;
   _57Y : ALIAS FOR I25[1].6;
   _5_LOWER_CROSS_BELT_HM : HOUR_METER := (HR_METER_DISPLAY := 2452, NEXT_SCHDL_MAINTENANCE := 2, MAINTENANCE_ALARM := 1);
   _5_LOWER_CROSS_BELT_RUNNING : BOOL;
   _5AUTO : ALIAS FOR B9[5].4;
   _5HAND : ALIAS FOR B9[5].3;
   _5M : ALIAS FOR O25[10].2;
   _5MB : ALIAS FOR B9[5].2;
   _5STB : ALIAS FOR B9[5].0;
   _5STPB : ALIAS FOR B9[5].1;
   _5Y : ALIAS FOR I25[2].2;
   _6AUTO : ALIAS FOR B9[6].4;
   _6HAND : ALIAS FOR B9[6].3;
   _6M : ALIAS FOR O25[10].3;
   _6MB : ALIAS FOR B9[6].2;
   _6STB : ALIAS FOR B9[6].0;
   _6STPB : ALIAS FOR B9[6].1;
   _6Y : ALIAS FOR I25[2].3;
   _700_AIR_GA : ALIAS FOR I8.3;
   _700_METER : ALIAS FOR I8.2;
   _700_PROBE : ALIAS FOR T22[9];
   _700_TREAT : ALIAS FOR I7.3;
   _700G_13_CL : ALIAS FOR B21[70].1;
   _700G_13_OP : ALIAS FOR B21[70].0;
   _700G_CLOSE : ALIAS FOR O12.9;
   _700G_OPEN : ALIAS FOR O12.8;
   _701_AIR_GA : ALIAS FOR I8.5;
   _701_FB : ALIAS FOR B21[1].3;
   _701_K_BYPA : ALIAS FOR I8.1;
   _701_K_TREA : ALIAS FOR I8.0;
   _701_METER : ALIAS FOR I8.4;
   _701_RB : ALIAS FOR B21[1].4;
   _701_REV_CN : ALIAS FOR C5[3];
   _701_STP : ALIAS FOR B21[1].2;
   _701_TRUCK_REVERSING_BELT_HM : HOUR_METER := (HR_METER_DISPLAY := 5981, NEXT_SCHDL_MAINTENANCE := 2, MAINTENANCE_ALARM := 1);
   _701_TRUCK_REVERSING_BELT_RUNNING : BOOL;
   _701F_HPB : ALIAS FOR B21[1].0;
   _701F_M : ALIAS FOR O25[10].11;
   _701F_OFF_T : ALIAS FOR T22[1];
   _701G_CLOSE : ALIAS FOR B21[71].13;
   _701G_OPEN : ALIAS FOR B21[71].12;
   _701K_GATE : ALIAS FOR B21[11].0;
   _701K_GATE1 : ALIAS FOR B21[11].1;
   _701K_GATE2 : ALIAS FOR B21[11].2;
   _701K_VALVE : ALIAS FOR O13.10;
   _701MR : ALIAS FOR O25[9].7;
   _701R_DELAY : ALIAS FOR T22[2];
   _701R_HPB : ALIAS FOR B21[1].1;
   _701Y : BOOL;
   _701YF : ALIAS FOR I25[2].11;
   _701YR : ALIAS FOR I25[1].7;
   _702_CLEAN_JUMP_BELT_HM : HOUR_METER := (HR_METER_DISPLAY := 3983, NEXT_SCHDL_MAINTENANCE := 2, MAINTENANCE_ALARM := 1);
   _702B : ALIAS FOR B21[2].2;
   _702H_START : ALIAS FOR B21[2].0;
   _702H_STOP : ALIAS FOR B21[2].1;
   _702M : ALIAS FOR O25[9].4;
   _702Y : ALIAS FOR I25[1].4;
   _703_TREATER_JUMP_BELT_HM : HOUR_METER := (HR_METER_DISPLAY := 2423, NEXT_SCHDL_MAINTENANCE := 2, MAINTENANCE_ALARM := 1);
   _703_TREATER_JUMP_BELT_RUNNING : BOOL;
   _703B : ALIAS FOR B21[3].2;
   _703H_START : ALIAS FOR B21[3].0;
   _703H_STOP : ALIAS FOR B21[3].1;
   _703M : ALIAS FOR O25[9].14;
   _703Y : ALIAS FOR I25[1].14;
   _704B : ALIAS FOR B21[4].2;
   _704H_START : ALIAS FOR B21[4].0;
   _704H_STOP : ALIAS FOR B21[4].1;
   _704M : ALIAS FOR O25[8].11;
   _704Y : ALIAS FOR I25[0].13;
   _705B : ALIAS FOR B21[5].2;
   _705H_START : ALIAS FOR B21[5].0;
   _705H_STOP : ALIAS FOR B21[5].1;
   _705M : ALIAS FOR O25[10].12;
   _705Y : ALIAS FOR I25[2].12;
   _705YA : ALIAS FOR I25[4].15;
   _706B : ALIAS FOR B21[6].2;
   _706H_START : ALIAS FOR B21[6].0;
   _706H_STOP : ALIAS FOR B21[6].1;
   _706M : ALIAS FOR O25[9].11;
   _706Y : ALIAS FOR I25[1].11;
   _707B : ALIAS FOR B21[7].2;
   _707M : ALIAS FOR O25[11].0;
   _707Y : ALIAS FOR I25[3].0;
   _708_BOT_CN : ALIAS FOR C5[5];
   _708G_BIN_1 : ALIAS FOR O9.15;
   _708G_BIN_2 : ALIAS FOR I7.4;
   _708G_CB13 : ALIAS FOR B21[8].0;
   _708G_CB131 : ALIAS FOR B21[8].1;
   _708G_CB132 : ALIAS FOR B21[8].2;
   _708G_HOLD : ALIAS FOR B21[8].3;
   _708G_HOLD1 : ALIAS FOR B21[8].6;
   _708G_RELEA : ALIAS FOR B21[8].4;
   _708G_RESET : ALIAS FOR B21[8].5;
   _709_BOT_CN : ALIAS FOR C5[6];
   _709G_BIN_1 : ALIAS FOR O10.15;
   _709G_BIN_2 : ALIAS FOR I7.5;
   _709G_CB19 : ALIAS FOR B21[9].0;
   _709G_CB191 : ALIAS FOR B21[9].1;
   _709G_CB192 : ALIAS FOR B21[9].2;
   _709G_HOLD : ALIAS FOR B21[9].3;
   _709G_HOLD1 : ALIAS FOR B21[9].6;
   _709G_RELEA : ALIAS FOR B21[9].4;
   _709G_RESET : ALIAS FOR B21[9].5;
   _709G_RUN_T : ALIAS FOR T22[8];
   _709G_TREAT : ALIAS FOR B21[9].7;
   _709G_TREAT1 : ALIAS FOR T22[10];
   _7AUTO : ALIAS FOR B9[7].4;
   _7HAND : ALIAS FOR B9[7].3;
   _7MB : ALIAS FOR B9[7].2;
   _7STB : ALIAS FOR B9[7].0;
   _7STPB : ALIAS FOR B9[7].1;
   _8AUTO : ALIAS FOR B9[8].4;
   _8HAND : ALIAS FOR B9[8].3;
   _8MB : ALIAS FOR B9[8].2;
   _8STB : ALIAS FOR B9[8].0;
   _8STPB : ALIAS FOR B9[8].1;
   _9_AIR_SV : ALIAS FOR O24[7].6;
   _9_BYPSS_GT : ALIAS FOR I24[6].1;
   _9_CAL_MOV : ALIAS FOR O24[7].2;
   _9_CAL_VALV : ALIAS FOR I24[6].5;
   _9_DRIP_GAT : ALIAS FOR O24[7].7;
   _9_GATE_SV : ALIAS FOR O24[7].0;
   _9_GATE_SV1 : ALIAS FOR O24[7].1;
   _9_SL_SW : ALIAS FOR B9[9].6;
   _9_SLW_SPEE : ALIAS FOR I25[3].12;
   _9_STP_SPEE : ALIAS FOR I25[3].13;
   _9_TREAT_MV : ALIAS FOR I24[6].6;
   _9_TREATER : ALIAS FOR I24[6].7;
   _9_TREATER_CONVAYOR_HM : HOUR_METER := (HR_METER_DISPLAY := 4578, NEXT_SCHDL_MAINTENANCE := 2, MAINTENANCE_ALARM := 1);
   _9_TREATER_CONVAYOR_RUNNING : BOOL;
   _9_TRT_M_ST : ALIAS FOR I24[6].3;
   _9_TRT_M_ST1 : ALIAS FOR I24[6].4;
   _9_TRT_MB : ALIAS FOR B3[9].0;
   _9_TRT_MOV : ALIAS FOR O24[7].4;
   _9_TRT_STB : ALIAS FOR B3[9].1;
   _9_TRT_STPB : ALIAS FOR B3[9].2;
   _9AUTO : ALIAS FOR B9[9].4;
   _9HAND : ALIAS FOR B9[9].3;
   _9M : ALIAS FOR O25[8].10;
   _9MB : ALIAS FOR B9[9].2;
   _9STB : ALIAS FOR B9[9].0;
   _9STPB : ALIAS FOR B9[9].1;
   _9Y : ALIAS FOR I25[0].10;
   _9YB : ALIAS FOR B9[9].5;
   A16 : INT[250] := ([24] := '0 ', [25] := '0 ', [26] := '0 ', [48] := '0 ', [110] := 'ge', [140] := 'ha', [150] := '10', [200] := 'cl', [210] := 'ov', [240] := 'le');
   A18 : INT[100] := ([13] := '9$00');
   A_ACC : ALIAS FOR N10[11];
   A_ACC_SEC : ALIAS FOR N10[13];
   A_HOLD_B : ALIAS FOR B3[1].4;
   A_HOLD_MB : ALIAS FOR B3[1].3;
   A_HOLD_REL : ALIAS FOR B3[1].5;
   A_MAIN_CNT : ALIAS FOR C5[0].PRE;
   A_MAIN_CNT1 : ALIAS FOR C5[0].ACC;
   A_MAIN_TRE : ALIAS FOR C5[0];
   A_PRESET : ALIAS FOR N10[10];
   A_PRESET_S : ALIAS FOR N10[12];
   A_RESET_PB : ALIAS FOR B3[1].2;
   A_SET : ALIAS FOR B3[1].6;
   A_STB_AUTO : ALIAS FOR B3[1].0;
   A_STPB_AUT : ALIAS FOR B3[1].1;
   A_TREATER : ALIAS FOR I24[6].8;
   A_TREATER1 : ALIAS FOR T4[59];
   ALARM_FIEL : ALIAS FOR T11[7];
   ALARM_HAND : ALIAS FOR B3[0].10;
   ALARM_HMI : ALIAS FOR B3[0].6;
   ALARM_HORN : ALIAS FOR O25[11].15;
   ALARM_HORN1 : ALIAS FOR O12.14;
   ALARM_INIT : ALIAS FOR B3[0].4;
   ALARM_LIGH : ALIAS FOR O13.15;
   ALARM_LT_O : ALIAS FOR T11[3];
   ALARM_SILE : ALIAS FOR I25[4].7;
   ALARM_SILE1 : ALIAS FOR I7.13;
   ALARM_SILE2 : ALIAS FOR B3[0].3;
   ALARM_SILE3 : ALIAS FOR B3[0].5;
   ALARM_SILE4 : ALIAS FOR B3[0].9;
   ALRM_LIGHT : ALIAS FOR O25[11].14;
   ALRM_SILEN : ALIAS FOR B3[0].7;
   Always_On : BOOL := 1;
   Analog : AI[160] := ([0].In := 104.0, [0].RawMin := 147.0, [0].RawMax := 16384.0, [0].EUMax := 3770.0, [1].In := 131.0, [1].RawMin := 147.0, [1].RawMax := 16384.0, [1].EUMax := 3770.0, [2].In := 1848.0, [2].RawMin := 1884.0, [2].RawMax := 16384.0, [2].EUMax := 4000.0, [20].In := 28816.0, [20].RawMin := 31000.0, [20].EUMax := 3200.0, [20].Out := 2974.5547, [21].In := 30336.0, [21].RawMax := 31000.0, [21].EUMax := 3200.0, [21].Out := 3131.458, [22].In := 30064.0, [22].RawMax := 31000.0, [22].EUMax := 3200.0, [22].Out := 3103.3806, [23].In := 7360.0, [23].RawMax := 31000.0, [23].EUMax := 3200.0, [23].Out := 759.74194, [24].In := 9136.0, [24].RawMax := 31000.0, [24].EUMax := 3200.0, [24].Out := 943.0709, [25].In := 28656.0, [25].RawMax := 31000.0, [25].EUMax := 3200.0, [25].Out := 2958.0386, [26].In := 28944.0, [26].RawMax := 31000.0, [26].EUMax := 3200.0, [26].Out := 2987.7676);
   B12 : DINT[100];
   B15 : DINT[100] := ([16] := 2#0000_0000_0000_0000_0000_0000_0000_0011, [17] := 2#0000_0000_0000_0000_0000_0000_0000_0011, [21] := 2#0000_0000_0000_0000_0000_0000_0000_0011, [22] := 2#0000_0000_0000_0000_0000_0000_0000_0011, [23] := 2#0000_0000_0000_0000_0000_0000_0000_0011, [30] := 2#0000_0000_0000_0000_0000_0000_0000_0011);
   B17 : DINT[30] := ([11] := 2#0000_0000_0000_0000_0000_0000_0000_0010, [12] := 2#0000_0000_0000_0000_0000_0000_0000_0111, [13] := 2#0000_0000_0000_0000_0000_0000_0000_0111, [14] := 2#0000_0000_0000_0000_0000_0000_0000_0010, [15] := 2#0000_0000_0000_0000_0000_0000_0000_0010, [16] := 2#0000_0000_0000_0000_0000_0000_0000_0111, [17] := 2#0000_0000_0000_0000_0000_0000_0000_0111, [21] := 2#0000_0000_0000_0000_0000_0000_0000_0010, [22] := 2#0000_0000_0000_0000_0000_0000_0000_0111, [23] := 2#0000_0000_0000_0000_0000_0000_0000_0111, [24] := 2#0000_0000_0000_0000_0000_0000_0000_0010, [25] := 2#0000_0000_0000_0000_0000_0000_0000_0111, [26] := 2#0000_0000_0000_0000_0000_0000_0000_0010);
   B183 : DINT[1] := ([0] := 2#0000_0000_0000_0000_0000_0000_0000_0001);
   B184 : DINT[1] := ([0] := 2#0000_0000_0000_0000_0000_0000_0000_0010);
   B194 : DINT[1];
   B204 : DINT[1];
   B21 : DINT[255];
   B214 : DINT[1];
   B224 : DINT[1] := ([0] := 2#0000_0000_0000_0000_0000_0000_0000_0010);
   B234 : DINT[1];
   B243 : DINT[1] := ([0] := 2#0000_0000_0000_0000_0000_0000_0000_0011);
   B244 : DINT[1] := ([0] := 2#0000_0000_0000_0000_0000_0000_0000_0010);
   B253 : DINT[100] := ([0] := 2#0000_0000_0000_0000_0000_0000_0000_0011);
   B254 : DINT[1] := ([0] := 2#0000_0000_0000_0000_0000_0000_0000_0010);
   B3 : DINT[250] := ([0] := 2#0000_0000_0000_0000_0000_0010_1011_0000, [101] := 2#0000_0000_0000_0000_0000_0000_0000_0010, [102] := 2#0000_0000_0000_0000_0000_0000_1000_0001);
   B9 : DINT[150] := ([1] := 2#0000_0000_0000_0000_0000_0000_0001_0100, [35] := 2#0000_0000_0000_0000_0000_0000_0001_0100, [42] := 2#0000_0000_0000_0000_0000_0000_0001_0100, [43] := 2#0000_0000_0000_0000_0000_0000_0011_0100, [45] := 2#0000_0000_0000_0000_0000_0000_0001_0100, [46] := 2#0000_0000_0000_0000_0000_0000_0001_0100, [48] := 2#0000_0000_0000_0000_0000_0000_0001_0100, [49] := 2#0000_0000_0000_0000_0000_0000_0001_0100, [50] := 2#0000_0000_0000_0000_0000_0000_0000_1000, [51] := 2#0000_0000_0000_0000_0000_0000_0001_0100, [52] := 2#0000_0000_0000_0000_0000_0000_0001_0100, [53] := 2#0000_0000_0000_0000_0000_0000_0001_0100, [54] := 2#0000_0000_0000_0000_0000_0000_0001_0100, [55] := 2#0000_0000_0000_0000_0000_0000_0001_0100, [57] := 2#0000_0000_0000_0000_0000_0000_0001_0100, [102] := 2#0000_0000_0000_0000_0000_0000_0000_1000, [103] := 2#0000_0000_0000_0000_0000_0000_0000_1000, [107] := 2#0000_0000_0000_0000_0000_0000_0011_0100, [108] := 2#0000_0000_0000_0000_0000_0000_0001_0100, [122] := 2#0000_0000_0000_0000_0000_0000_0001_0100, [123] := 2#0000_0000_0000_0000_0000_0000_0001_0100);
   Beta : BOOL := 1;
   BIN_1_CLOSE : BOOL;
   BIN_1_OPEN : BOOL;
   BIN_2_CLOSE : BOOL;
   BIN_2_OPEN : BOOL;
   BIN_3_CLOSE : BOOL;
   BIN_3_OPEN : BOOL;
   BIN_4_CLOSE : BOOL;
   BIN_4_OPEN : BOOL;
   BIN_5_CLOSE : BOOL;
   BIN_5_OPEN : BOOL;
   BIN_6_CLOSE : BOOL;
   BIN_6_OPEN : BOOL;
   BIN_7_CLOSE : BOOL;
   BIN_7_OPEN : BOOL;
   Bin_Config : BOOL := 1;
   C5 : COUNTER[50] := ([0].PRE := 3000, [1].ACC := 5, [1].DN := 1, [2].PRE := 3000, [3].PRE := 2, [4].PRE := 400000, [5].PRE := 5000, [5].CU := 1, [6].PRE := 9999, [6].CU := 1, [11].PRE := 1200, [12].PRE := 30, [13].PRE := 3000, [14].PRE := 36, [15].PRE := 1500, [16].PRE := 3000, [17].PRE := 3000, [21].PRE := 3000, [22].PRE := 3000, [23].PRE := 3000, [24].PRE := 3000, [25].PRE := 3000, [26].PRE := 3000, [27].CU := 1, [28].CU := 1, [29].CU := 1, [30].PRE := 20000, [32].PRE := 20000, [33].PRE := 20000, [34].PRE := 20000, [35].PRE := 20000, [36].PRE := 20000, [37].PRE := 20000, [38].PRE := 20000, [39].PRE := 20000);
   CAL_K_FACT : ALIAS FOR F8[0];
   CAL_RESET : ALIAS FOR B15[50].0;
   Calibration_Max : REAL := 4000.0;
   CG13_METR : ALIAS FOR I8.15;
   CG_13_AIR : ALIAS FOR I8.13;
   CG_19_AIR : ALIAS FOR I8.12;
   CG_19_METR : ALIAS FOR I8.14;
   CHEM_PUMP_1 : STRING := 'water';
   CHEM_PUMP_10 : STRING := 'oil';
   CHEM_PUMP_11 : STRING := 'apron';
   CHEM_PUMP_12 : STRING := 'stamina';
   CHEM_PUMP_13 : STRING := 'TEST13';
   CHEM_PUMP_14 : STRING := 'oil';
   CHEM_PUMP_15 : STRING := 'red';
   CHEM_PUMP_2 : STRING := 'alba red';
   CHEM_PUMP_3 : STRING := 'evergol';
   CHEM_PUMP_4 : STRING := 'macho';
   CHEM_PUMP_5 : STRING := 'vib ex';
   CHEM_PUMP_6 : STRING := 'bio st';
   CHEM_PUMP_7 : STRING := 'tbz';
   CHEM_PUMP_8 : STRING := 'wuxal';
   CHEM_PUMP_9 : STRING := 'BLUE';
   CIMBRA_BIN : ALIAS FOR I25[3].10;
   CIMBRIA_BI : ALIAS FOR B15[30].0;
   CIMBRIA_BI1 : ALIAS FOR B15[30].1;
   CIMBRIA_BIN_EMPTY : BOOL;
   CIMBRIA_BIN_FULL : BOOL;
   CIMBRIA_FAN_ON : BOOL := 1;
   CIMBRIA_FAN_SPD_INPUT : DINT := 30;
   CIMBRIA_HI : ALIAS FOR B15[30].2;
   CIMBRIA_OUTPUT_SPD : DINT := 30;
   Cleaning_Motors : udt_Motor[100] := ([0].Motor_Control.Motor_Amps := 1.3896561, [1].Motor_Control.Motor_Amps := 1.006918, [2].Motor_Control.Motor_Amps := 0.8792738, [3].Motor_Control.Motor_Amps := 2.5666564);
   CLR_SORT_ASP_DELAY : TIMER := (PRE := 5000, ACC := 5002, EN := 1, DN := 1);
   CLR_SORT_ASPBLR_DELAY : TIMER := (PRE := 5000, ACC := 5004, EN := 1, DN := 1);
   CLR_SORT_LEG_DELAY : TIMER := (PRE := 5000, ACC := 5003, EN := 1, DN := 1);
   CLR_SORT_LEG_SPD10 : ALIAS FOR Local:0:I.Data.3;
   CLR_SORT_LEG_SPD20 : ALIAS FOR Local:0:I.Data.4;
   CONC13_COL : ALIAS FOR N7[93];
   CONC13_OP : ALIAS FOR A18[3];
   CONC13_PUM : ALIAS FOR N7[83];
   CONC13_SET : ALIAS FOR A18[0];
   CONC13_SET1 : ALIAS FOR B21[8].14;
   CONC19_COL : ALIAS FOR N7[99];
   CONC19_OP : ALIAS FOR A18[13];
   CONC19_PUM : ALIAS FOR N7[89];
   CONC19_SET : ALIAS FOR B21[9].14;
   CONC_13_NO : ALIAS FOR B21[8].15;
   CONC_19_NO : ALIAS FOR B21[9].15;
   CONC_19_SE : ALIAS FOR A18[10];
   ConcretePlantIn : DINT := 2;
   ConcretePlantOut : DINT := 1; {produced}
   Config_Save_Binss : BOOL;
   ConfigureVariety : Variety;
   Consumed : DINT;
   CP_Remote_Air_Gate_On : DINT; {produced}
   CP_Remote_Air_Gate_Open_In : DINT;
   CP_Remote_Andco_Auto_In : DINT;
   CP_Remote_Andoc_Out : udt_Andco_Remote_Out[32]; {produced}
   CP_Remote_Belt_In : udt_Motor_Remote_In[10] := ([1].Spd_10_Out := 1, [1].Amps := -0.32500002, [2].Spd_10_Out := 1, [2].Amps := -0.425, [3].Spd_10_Out := 1, [3].Amps := -0.5125);
   CP_Remote_Belt_Start : DINT; {produced}
   CP_Remote_Leg_In : udt_Motor_Remote_In := (Spd_20_Out := 1, Spd_10_Out := 1, Amps := -0.22500001);
   CP_Remote_Leg_Start : DINT; {produced}
   cpBinGateRates : DINT[50] := ([1] := 73, [3] := 180, [5] := 531, [7] := 117, [10] := 147, [13] := 269, [19] := 173);
   cpBINOPEN : DINT;
   cpCleanBulk : BOOL;
   cpTicketBinActive : DINT;
   cpTicketBinSet : DINT;
   cpVAR_BINARRAY : STRING[50] := ([1] := '823019-Diva Spring-Certified-WSU -SWW Seed Wheat', [3] := '823007-WB 6121 spring-Certified - Monsanto  - SWW Seed Wheat', [4] := 'reg duet', [5] := '823001-ArtDeco-Certified-Limagrain -SWW Seed Wheat', [10] := '823007-WB 6121 spring-Certified-Monsanto -SWW Seed Wheat', [11] := '823014-Skiles-Certified-OSU -SWW Seed Wheat', [20] := '823010-Bobtail-Certified-OSU -SWW Seed Wheat');
   cpVAR_CNT_ONS : DINT;
   cpVarTrimTemp : STRING := '823026';
   Dev : DINT := 6145; {produced}
   DIST_MOVE : ALIAS FOR I3.10;
   DIST_TO_CL : ALIAS FOR I7.2;
   DS_CLEAN_B : ALIAS FOR O13.5;
   DS_DLY_OFF : ALIAS FOR T4[33];
   DS_M : ALIAS FOR O24[1].0;
   DS_M_B : ALIAS FOR B3[101].0;
   DS_MOV_CCW : ALIAS FOR B3[100].13;
   DS_MOV_CW : ALIAS FOR B3[100].12;
   DS_MOVE_SE : ALIAS FOR T4[32];
   DS_POS8 : ALIAS FOR O13.7;
   DS_POS9 : ALIAS FOR O13.8;
   DS_POS_1 : ALIAS FOR I24[0].2;
   DS_POS_10 : ALIAS FOR I24[0].11;
   DS_POS_11 : ALIAS FOR B3[100].11;
   DS_POS_1_B : ALIAS FOR B3[100].2;
   DS_POS_2 : ALIAS FOR I24[0].3;
   DS_POS_2_B : ALIAS FOR B3[100].3;
   DS_POS_3 : ALIAS FOR I24[0].4;
   DS_POS_3_B : ALIAS FOR B3[100].4;
   DS_POS_4 : ALIAS FOR I24[0].5;
   DS_POS_4_B : ALIAS FOR B3[100].5;
   DS_POS_5 : ALIAS FOR I24[0].6;
   DS_POS_5_B : ALIAS FOR B3[100].6;
   DS_POS_6 : ALIAS FOR I24[0].7;
   DS_POS_6_B : ALIAS FOR B3[100].7;
   DS_POS_7 : ALIAS FOR I24[0].8;
   DS_POS_7_B : ALIAS FOR B3[100].8;
   DS_POS_8 : ALIAS FOR I24[0].9;
   DS_POS_8_B : ALIAS FOR B3[100].9;
   DS_POS_9 : ALIAS FOR I24[0].10;
   DS_POS_9_B : ALIAS FOR B3[100].10;
   DS_SEEK_1 : ALIAS FOR B3[102].1;
   DS_SEEK_10 : ALIAS FOR B3[102].10;
   DS_SEEK_2 : ALIAS FOR B3[102].2;
   DS_SEEK_3 : ALIAS FOR B3[102].3;
   DS_SEEK_4 : ALIAS FOR B3[102].4;
   DS_SEEK_5 : ALIAS FOR B3[102].5;
   DS_SEEK_6 : ALIAS FOR B3[102].6;
   DS_SEEK_7 : ALIAS FOR B3[102].7;
   DS_SEEK_8 : ALIAS FOR B3[102].8;
   DS_SEEK_9 : ALIAS FOR B3[102].9;
   DS_SET_IN : ALIAS FOR N10[0];
   DS_SP_UP_B : ALIAS FOR B3[100].0;
   DS_SPOUT_C : ALIAS FOR O24[1].3;
   DS_SPOUT_C1 : ALIAS FOR O24[1].4;
   DS_SPOUT_C2 : ALIAS FOR B3[101].3;
   DS_SPOUT_C3 : ALIAS FOR B3[101].4;
   DS_SPOUT_D : ALIAS FOR I24[0].1;
   DS_SPOUT_D1 : ALIAS FOR O24[1].1;
   DS_SPOUT_D2 : ALIAS FOR B3[100].1;
   DS_SPOUT_D3 : ALIAS FOR B3[101].1;
   DS_SPOUT_U : ALIAS FOR I24[0].0;
   DS_SPOUT_U1 : ALIAS FOR O24[1].2;
   DS_SPOUT_U2 : ALIAS FOR B3[101].2;
   DS_START_M : ALIAS FOR B3[102].11;
   DS_STOP_MO : ALIAS FOR B3[102].0;
   DS_T21 : ALIAS FOR O13.0;
   DS_T22 : ALIAS FOR O13.1;
   DS_T23 : ALIAS FOR O13.9;
   DS_T231 : ALIAS FOR O13.2;
   DS_T24 : ALIAS FOR O13.3;
   DS_T25 : ALIAS FOR O13.4;
   DS_T26 : ALIAS FOR O13.6;
   F8 : REAL[27] := ([0] := 1.2, [1] := 1.0, [2] := 14748.0, [3] := 1.0, [4] := 15440.0, [5] := 1.0, [6] := 14244.0, [7] := 1.0, [8] := 13454.0, [9] := 1.0, [10] := 14460.0, [11] := 1.0, [12] := 6343.0, [13] := 1.0, [14] := 8758.0, [15] := 1.0, [16] := 15944.0, [17] := 1.0, [18] := 15184.0, [19] := 1.0, [20] := 15741.0, [21] := 1.0, [22] := 15276.0, [23] := 1.0, [24] := 14611.0, [25] := 1.0, [26] := 15145.0);
   Gates : STRING;
   hCLR_SORT_LEG_SPD10 : BOOL := 1;
   hCLR_SORT_LEG_SPD20 : BOOL := 1;
   hCLR_SORT_STB : BOOL;
   hCLR_SORT_STRT : BOOL;
   hN_RECVING_PIT_GATE_CLSPB : BOOL;
   hN_RECVING_PIT_GATE_OPNPB : BOOL;
   hSURGE_BIN_HI : BOOL;
   hSURGE_BIN_LO : BOOL;
   I1 : ALIAS FOR R1S0_AENTR:1:I.Data;
   I16 : INT[16] := ([0] := 2#0011_1001_1001_1100, [1] := 2#0011_1100_0101_0000, [2] := 2#0011_0111_1010_0100, [3] := 2#0011_0100_1000_1110, [4] := 2#0011_1000_0111_1100, [5] := 2#0001_1000_1100_0111, [6] := 2#0010_0010_0011_0110, [7] := 2#0011_1110_0100_1000, [8] := 2#0000_1000_0101_1010, [9] := 2#0000_1000_0101_1010, [10] := 2#0000_1000_0101_1010, [11] := 2#0000_1000_0101_1010, [12] := 2#0000_1000_0101_1010, [13] := 2#0000_1000_0101_1010, [14] := 2#0000_1000_0101_1010, [15] := 2#0000_1000_0101_1010);
   I16_0 : ALIAS FOR N20[0];
   I16_000 : ALIAS FOR I16[0];
   I16_001 : ALIAS FOR I16[1];
   I16_002 : ALIAS FOR I16[2];
   I16_003 : ALIAS FOR I16[3];
   I16_004 : ALIAS FOR I16[4];
   I16_005 : ALIAS FOR I16[5];
   I16_006 : ALIAS FOR I16[6];
   I16_007 : ALIAS FOR I16[7];
   I16_1 : ALIAS FOR N20[1];
   I16_2 : ALIAS FOR N20[2];
   I16_3 : ALIAS FOR N20[3];
   I16_4 : ALIAS FOR N20[4];
   I16_5 : ALIAS FOR N20[5];
   I16_6 : ALIAS FOR N20[6];
   I16_7 : ALIAS FOR N20[7];
   I17 : INT[16] := ([0] := 2#0011_1011_0101_0000, [1] := 2#0011_1101_0111_1101, [2] := 2#0011_1011_1010_1111, [3] := 2#0011_1001_0001_0011, [4] := 2#0011_1011_0010_1001, [5] := 2#0001_1100_1010_0101, [6] := 2#0001_1100_1010_1111, [7] := 2#0001_1100_1010_0010, [8] := 2#0000_1000_0101_1010, [9] := 2#0000_1000_0101_1010, [10] := 2#0000_1000_0101_1010, [11] := 2#0000_1000_0101_1010, [12] := 2#0000_1000_0101_1010, [13] := 2#0000_1000_0101_1010, [14] := 2#0000_1000_0101_1010, [15] := 2#0000_1000_0101_1010);
   I17_000 : ALIAS FOR I17[0];
   I17_001 : ALIAS FOR I17[1];
   I17_002 : ALIAS FOR I17[2];
   I17_003 : ALIAS FOR I17[3];
   I17_004 : ALIAS FOR I17[4];
   I17_005 : ALIAS FOR I17[5];
   I17_006 : ALIAS FOR I17[6];
   I17_007 : ALIAS FOR I17[7];
   I18 : INT[16] := ([0] := 2#0000_0101_0101_0011, [1] := 2#0000_0111_0011_1000, [2] := 2#0000_0000_1000_0011, [3] := 2#0000_0000_0110_1000, [4] := 2#0000_0111_0111_1100, [5] := 2#0000_0111_0110_0101, [6] := 2#0000_1100_1100_1101, [7] := 2#0000_1100_1100_1101, [8] := 2#0000_1000_0101_1010, [9] := 2#0000_1000_0101_1010, [10] := 2#0000_1000_0101_1010, [11] := 2#0000_1000_0101_1010, [12] := 2#0000_1000_0101_1010, [13] := 2#0000_1000_0101_1010, [14] := 2#0001_1010_1001_1101, [15] := 2#0001_1010_1001_1101);
   I18_000 : ALIAS FOR I18[0];
   I18_001 : ALIAS FOR I18[1];
   I18_002 : ALIAS FOR I18[2];
   I18_003 : ALIAS FOR I18[3];
   I18_007 : ALIAS FOR I18[7];
   I1_000_Bit00 : ALIAS FOR I1.0;
   I1_000_Bit01 : ALIAS FOR I1.1;
   I1_000_Bit02 : ALIAS FOR I1.2;
   I1_000_Bit03 : ALIAS FOR I1.3;
   I1_000_Bit04 : ALIAS FOR I1.4;
   I1_000_Bit05 : ALIAS FOR I1.5;
   I1_000_Bit06 : ALIAS FOR I1.6;
   I1_000_Bit07 : ALIAS FOR I1.7;
   I1_000_Bit08 : ALIAS FOR I1.8;
   I1_000_Bit09 : ALIAS FOR I1.9;
   I1_000_Bit10 : ALIAS FOR I1.10;
   I1_000_Bit11 : ALIAS FOR I1.11;
   I1_000_Bit12 : ALIAS FOR I1.12;
   I1_000_Bit13 : ALIAS FOR I1.13;
   I1_000_Bit14 : ALIAS FOR I1.14;
   I1_000_Bit15 : ALIAS FOR I1.15;
   I2 : ALIAS FOR R1S0_AENTR:2:I.Data;
   I24 : INT[32] := ([0] := 2#0000_0001_0000_0010, [6] := 2#0010_0000_1000_0110, [7] := 2#0010_0000_1000_0110);
   I24_000_Bit00 : ALIAS FOR I24[0].0;
   I24_000_Bit01 : ALIAS FOR I24[0].1;
   I24_000_Bit02 : ALIAS FOR I24[0].2;
   I24_000_Bit03 : ALIAS FOR I24[0].3;
   I24_000_Bit04 : ALIAS FOR I24[0].4;
   I24_000_Bit05 : ALIAS FOR I24[0].5;
   I24_000_Bit06 : ALIAS FOR I24[0].6;
   I24_000_Bit07 : ALIAS FOR I24[0].7;
   I24_000_Bit08 : ALIAS FOR I24[0].8;
   I24_000_Bit09 : ALIAS FOR I24[0].9;
   I24_000_Bit10 : ALIAS FOR I24[0].10;
   I24_000_Bit11 : ALIAS FOR I24[0].11;
   I24_004_Bit00 : ALIAS FOR I24[4].0;
   I24_004_Bit01 : ALIAS FOR I24[4].1;
   I24_004_Bit02 : ALIAS FOR I24[4].2;
   I24_004_Bit03 : ALIAS FOR I24[4].3;
   I24_004_Bit04 : ALIAS FOR I24[4].4;
   I24_004_Bit05 : ALIAS FOR I24[4].5;
   I24_004_Bit06 : ALIAS FOR I24[4].6;
   I24_004_Bit07 : ALIAS FOR I24[4].7;
   I24_004_Bit08 : ALIAS FOR I24[4].8;
   I24_004_Bit09 : ALIAS FOR I24[4].9;
   I24_004_Bit10 : ALIAS FOR I24[4].10;
   I24_004_Bit11 : ALIAS FOR I24[4].11;
   I24_004_Bit12 : ALIAS FOR I24[4].12;
   I24_006_Bit01 : ALIAS FOR I24[6].1;
   I24_006_Bit02 : ALIAS FOR I24[6].2;
   I24_006_Bit07 : ALIAS FOR I24[6].7;
   I24_006_Bit08 : ALIAS FOR I24[6].8;
   I24_006_Bit13 : ALIAS FOR I24[6].13;
   I24_021_Bit00 : ALIAS FOR I24[21].0;
   I24_021_Bit01 : ALIAS FOR I24[21].1;
   I24_021_Bit02 : ALIAS FOR I24[21].2;
   I24_021_Bit03 : ALIAS FOR I24[21].3;
   I24_021_Bit04 : ALIAS FOR I24[21].4;
   I24_021_Bit05 : ALIAS FOR I24[21].5;
   I24_021_Bit06 : ALIAS FOR I24[21].6;
   I24_021_Bit07 : ALIAS FOR I24[21].7;
   I24_021_Bit08 : ALIAS FOR I24[21].8;
   I25 : INT[32] := ([0] := 2#0101_0011_1101_1110, [1] := 2#0011_0011_0100_0010, [2] := 2#1110_0000_0100_0000, [3] := 2#1101_0000_0000_1010, [4] := 2#0110_0000_0000_1101);
   I25_000_Bit00 : ALIAS FOR I25[0].0;
   I25_000_Bit01 : ALIAS FOR I25[0].1;
   I25_000_Bit02 : ALIAS FOR I25[0].2;
   I25_000_Bit03 : ALIAS FOR I25[0].3;
   I25_000_Bit04 : ALIAS FOR I25[0].4;
   I25_000_Bit06 : ALIAS FOR I25[0].6;
   I25_000_Bit07 : ALIAS FOR I25[0].7;
   I25_000_Bit08 : ALIAS FOR I25[0].8;
   I25_000_Bit09 : ALIAS FOR I25[0].9;
   I25_000_Bit10 : ALIAS FOR I25[0].10;
   I25_000_Bit12 : ALIAS FOR I25[0].12;
   I25_000_Bit13 : ALIAS FOR I25[0].13;
   I25_000_Bit14 : ALIAS FOR I25[0].14;
   I25_000_Bit15 : ALIAS FOR I25[0].15;
   I25_001_Bit00 : ALIAS FOR I25[1].0;
   I25_001_Bit01 : ALIAS FOR I25[1].1;
   I25_001_Bit02 : ALIAS FOR I25[1].2;
   I25_001_Bit03 : ALIAS FOR I25[1].3;
   I25_001_Bit04 : ALIAS FOR I25[1].4;
   I25_001_Bit05 : ALIAS FOR I25[1].5;
   I25_001_Bit06 : ALIAS FOR I25[1].6;
   I25_001_Bit07 : ALIAS FOR I25[1].7;
   I25_001_Bit08 : ALIAS FOR I25[1].8;
   I25_001_Bit09 : ALIAS FOR I25[1].9;
   I25_001_Bit10 : ALIAS FOR I25[1].10;
   I25_001_Bit11 : ALIAS FOR I25[1].11;
   I25_001_Bit12 : ALIAS FOR I25[1].12;
   I25_001_Bit13 : ALIAS FOR I25[1].13;
   I25_001_Bit14 : ALIAS FOR I25[1].14;
   I25_001_Bit15 : ALIAS FOR I25[1].15;
   I25_002_Bit00 : ALIAS FOR I25[2].0;
   I25_002_Bit01 : ALIAS FOR I25[2].1;
   I25_002_Bit02 : ALIAS FOR I25[2].2;
   I25_002_Bit03 : ALIAS FOR I25[2].3;
   I25_002_Bit04 : ALIAS FOR I25[2].4;
   I25_002_Bit05 : ALIAS FOR I25[2].5;
   I25_002_Bit06 : ALIAS FOR I25[2].6;
   I25_002_Bit08 : ALIAS FOR I25[2].8;
   I25_002_Bit09 : ALIAS FOR I25[2].9;
   I25_002_Bit10 : ALIAS FOR I25[2].10;
   I25_002_Bit11 : ALIAS FOR I25[2].11;
   I25_002_Bit12 : ALIAS FOR I25[2].12;
   I25_002_Bit13 : ALIAS FOR I25[2].13;
   I25_002_Bit14 : ALIAS FOR I25[2].14;
   I25_002_Bit15 : ALIAS FOR I25[2].15;
   I25_003_Bit00 : ALIAS FOR I25[3].0;
   I25_003_Bit01 : ALIAS FOR I25[3].1;
   I25_003_Bit03 : ALIAS FOR I25[3].3;
   I25_003_Bit10 : ALIAS FOR I25[3].10;
   I25_003_Bit12 : ALIAS FOR I25[3].12;
   I25_003_Bit13 : ALIAS FOR I25[3].13;
   I25_003_Bit14 : ALIAS FOR I25[3].14;
   I25_003_Bit15 : ALIAS FOR I25[3].15;
   I25_004_Bit00 : ALIAS FOR I25[4].0;
   I25_004_Bit01 : ALIAS FOR I25[4].1;
   I25_004_Bit02 : ALIAS FOR I25[4].2;
   I25_004_Bit03 : ALIAS FOR I25[4].3;
   I25_004_Bit06 : ALIAS FOR I25[4].6;
   I25_004_Bit07 : ALIAS FOR I25[4].7;
   I25_004_Bit14 : ALIAS FOR I25[4].14;
   I2_000_Bit00 : ALIAS FOR I2.0;
   I2_000_Bit02 : ALIAS FOR I2.2;
   I2_000_Bit03 : ALIAS FOR I2.3;
   I2_000_Bit05 : ALIAS FOR I2.5;
   I2_000_Bit06 : ALIAS FOR I2.6;
   I2_000_Bit07 : ALIAS FOR I2.7;
   I2_000_Bit08 : ALIAS FOR I2.8;
   I2_000_Bit09 : ALIAS FOR I2.9;
   I2_000_Bit10 : ALIAS FOR I2.10;
   I2_000_Bit11 : ALIAS FOR I2.11;
   I2_000_Bit12 : ALIAS FOR I2.12;
   I2_000_Bit13 : ALIAS FOR I2.13;
   I2_000_Bit14 : ALIAS FOR I2.14;
   I3 : ALIAS FOR R1S0_AENTR:3:I.Data;
   I3_000_Bit00 : ALIAS FOR I3.0;
   I3_000_Bit01 : ALIAS FOR I3.1;
   I3_000_Bit02 : ALIAS FOR I3.2;
   I3_000_Bit03 : ALIAS FOR I3.3;
   I3_000_Bit04 : ALIAS FOR I3.4;
   I3_000_Bit05 : ALIAS FOR I3.5;
   I3_000_Bit06 : ALIAS FOR I3.6;
   I3_000_Bit07 : ALIAS FOR I3.7;
   I3_000_Bit08 : ALIAS FOR I3.8;
   I3_000_Bit09 : ALIAS FOR I3.9;
   I3_000_Bit10 : ALIAS FOR I3.10;
   I3_000_Bit11 : ALIAS FOR I3.11;
   I3_000_Bit12 : ALIAS FOR I3.12;
   I3_000_Bit14 : ALIAS FOR I3.14;
   I4 : ALIAS FOR R1S0_AENTR:4:I.Data;
   I4_000_Bit00 : ALIAS FOR I4.0;
   I4_000_Bit02 : ALIAS FOR I4.2;
   I4_000_Bit04 : ALIAS FOR I4.4;
   I4_000_Bit09 : ALIAS FOR I4.9;
   I4_000_Bit10 : ALIAS FOR I4.10;
   I4_000_Bit11 : ALIAS FOR I4.11;
   I4_000_Bit12 : ALIAS FOR I4.12;
   I4_000_Bit13 : ALIAS FOR I4.13;
   I4_000_Bit14 : ALIAS FOR I4.14;
   I4_000_Bit15 : ALIAS FOR I4.15;
   I5 : ALIAS FOR R1S0_AENTR:5:I.Data;
   I6 : ALIAS FOR R1S0_AENTR:6:I.Data;
   I7 : ALIAS FOR R1S0_AENTR:7:I.Data;
   I7_000_Bit02 : ALIAS FOR I7.2;
   I7_000_Bit03 : ALIAS FOR I7.3;
   I7_000_Bit04 : ALIAS FOR I7.4;
   I7_000_Bit05 : ALIAS FOR I7.5;
   I7_000_Bit13 : ALIAS FOR I7.13;
   I7_000_Bit14 : ALIAS FOR I7.14;
   I7_000_Bit15 : ALIAS FOR I7.15;
   I8 : ALIAS FOR R1S0_AENTR:8:I.Data;
   I8_000_Bit00 : ALIAS FOR I8.0;
   I8_000_Bit02 : ALIAS FOR I8.2;
   I8_000_Bit03 : ALIAS FOR I8.3;
   I8_000_Bit04 : ALIAS FOR I8.4;
   I8_000_Bit05 : ALIAS FOR I8.5;
   I8_000_Bit06 : ALIAS FOR I8.6;
   I8_000_Bit07 : ALIAS FOR I8.7;
   I8_000_Bit08 : ALIAS FOR I8.8;
   I8_000_Bit09 : ALIAS FOR I8.9;
   I8_000_Bit10 : ALIAS FOR I8.10;
   I8_000_Bit11 : ALIAS FOR I8.11;
   I8_000_Bit12 : ALIAS FOR I8.12;
   IE8_BTR_FL : ALIAS FOR N23[0];
   indexTbl : DINT;
   indexTblOld : DINT;
   indexTRTTbl : DINT;
   InEUMax : REAL;
   K_FACTOR : ALIAS FOR N14[80];
   M0_24 : INT[3300] := ([100] := -32640, [200] := -32768, [300] := 128, [400] := -32768, [500] := -32640, [700] := -32640, [800] := -32768, [900] := -32640);
   M0_25 : INT[3300] := ([100] := -32640, [300] := -32640, [500] := 128, [600] := -32768);
   M1_24 : INT[3300];
   M1_25 : INT[3300];
   M701_SLOW : ALIAS FOR I8.6;
   M701_STOP : ALIAS FOR I8.7;
   M702_SLOW : ALIAS FOR I8.8;
   M702_STOP : ALIAS FOR I8.9;
   M703_SLOW : ALIAS FOR I8.10;
   M703_STOP : ALIAS FOR I8.11;
   MAIN_TIMER : ALIAS FOR T11[0];
   MAIN_TIMER1 : ALIAS FOR T11[1];
   MASTER_FAU : ALIAS FOR B3[0].1;
   MASTER_STO : ALIAS FOR B3[0].2;
   MTR_125_RUNNING : ALIAS FOR Local:0:I.Data.11;
   MTR_125MB : ALIAS FOR Local:5:O.Data.0;
   MTR_126_RUNNING : ALIAS FOR Local:0:I.Data.6;
   MTR_126M : ALIAS FOR Local:5:O.Data.1;
   MTR_126MB : BOOL := 1;
   MTR_127_RUNNING : ALIAS FOR Local:0:I.Data.7;
   MTR_127M : ALIAS FOR Local:5:O.Data.2;
   MTR_127MB : BOOL := 1;
   MTR_128_RUNNING : ALIAS FOR Local:0:I.Data.5;
   MTR_128M : ALIAS FOR Local:5:O.Data.3;
   MTR_128MB : BOOL := 1;
   N10 : DINT[30] := ([0] := 7, [1] := 7, [10] := 500, [12] := 3000);
   N13 : DINT[100] := ([4] := 80, [14] := 43, [24] := 35, [34] := 30, [44] := 29, [54] := 30, [64] := 30, [74] := 40, [84] := 22);
   N14 : DINT[84] := ([11] := 3173, [12] := 3523, [13] := 2924, [14] := 3485, [15] := 3442, [16] := 1402, [17] := 2895, [21] := 3209, [22] := 3053, [23] := 3621, [24] := 3332, [25] := 4010, [26] := 3739, [31] := 1, [32] := 7589, [33] := 7589, [34] := 1, [35] := 9417, [36] := 9417, [37] := 1, [38] := 10027, [39] := 10027, [40] := 1, [41] := 8, [43] := 1, [44] := 8771, [45] := 8771, [46] := 1, [47] := 8060, [48] := 8060, [49] := 1, [50] := 6101, [51] := 6101, [52] := 1, [53] := 15066, [54] := 15066, [55] := 1, [56] := 10230, [57] := 10230, [58] := 1, [59] := 9011, [60] := 9011, [61] := 1, [62] := 9440, [63] := 9440, [64] := 1, [65] := 7454, [66] := 7454, [67] := 1, [68] := 9863, [69] := 9863, [80] := 120);
   N180 : DINT[68] := ([0] := 160, [1] := 14932, [2] := 27374, [3] := 14300, [4] := 23411, [5] := 12, [7] := 3026, [8] := 239, [10] := -256, [50] := 128, [51] := 9, [52] := 220, [54] := 1, [55] := 220, [60] := 25600, [61] := 9, [62] := 220, [64] := 1024, [66] := 220);
   N181 : DINT[1];
   N182 : DINT[2] := ([0] := -9, [1] := -9);
   N190 : DINT[68] := ([0] := 14, [10] := 23340, [14] := 15, [15] := 3840, [50] := -32640, [51] := 1, [52] := 210, [54] := 14, [55] := 210, [61] := 1, [62] := 210, [64] := 25600, [65] := 14, [66] := 210);
   N191 : DINT[1];
   N192 : DINT[2] := ([0] := -9, [1] := -9);
   N193 : DINT[1] := ([0] := 9);
   N20 : DINT[30] := ([0] := 2138, [1] := 2138, [2] := 2138, [3] := 2138, [4] := 2138, [5] := 2138, [6] := 2138, [7] := 2138, [10] := 2138, [11] := 2138, [12] := 2138, [13] := 2138, [14] := 2138, [15] := 2138, [16] := 2138, [17] := 2138, [20] := 2138, [21] := 2138, [22] := 2138, [23] := 2138, [24] := 2138, [25] := 2138, [26] := 2717, [27] := 2717);
   N200 : DINT[68] := ([10] := 400, [11] := 24800, [12] := 27383, [13] := 23767, [14] := 15, [15] := 3840, [50] := -32640, [51] := 1, [52] := 200, [54] := 14, [55] := 200, [61] := 1, [62] := 200, [64] := 25600, [65] := 14, [66] := 200);
   N201 : DINT[1];
   N202 : DINT[2] := ([0] := -9, [1] := -9);
   N203 : DINT[1] := ([0] := 9);
   N210 : DINT[68] := ([0] := 14, [10] := 7040, [11] := 2, [14] := 15, [15] := 3840, [50] := -32640, [51] := 1, [52] := 240, [54] := 14, [55] := 240, [60] := 1024, [62] := 240, [64] := 25600, [65] := 14, [66] := 240);
   N211 : DINT[1];
   N212 : DINT[2] := ([0] := -9, [1] := -9);
   N213 : DINT[1] := ([0] := 9);
   N220 : DINT[68] := ([10] := 9280, [11] := 9600, [12] := 9600, [13] := 12800, [14] := 15, [15] := 3840, [50] := -32640, [51] := 1, [52] := 230, [54] := 14, [55] := 230, [61] := 1, [62] := 230, [64] := 1024, [66] := 230);
   N221 : DINT[1];
   N222 : DINT[2] := ([0] := -9, [1] := -9);
   N223 : DINT[1] := ([0] := 3);
   N23 : DINT[5] := ([0] := 11, [1] := 60, [2] := 11, [3] := 60);
   N230 : DINT[68] := ([10] := 24720, [11] := 13760, [12] := 11200, [13] := 9600, [14] := 15, [15] := 3840, [50] := -32640, [51] := 1, [52] := 220, [54] := 14, [55] := 220, [61] := 1, [62] := 220, [64] := 25600, [65] := 14, [66] := 220);
   N231 : DINT[1];
   N232 : DINT[2] := ([0] := -9, [1] := -9);
   N233 : DINT[1] := ([0] := 9);
   N24 : DINT[31] := ([0] := 100, [1] := 1, [2] := 100, [3] := 1, [4] := 5, [5] := 5, [6] := 60, [7] := 1, [8] := 100, [9] := 1, [10] := 100, [11] := 1, [12] := 5, [13] := 5, [14] := 60, [15] := 1);
   N240 : DINT[68] := ([8] := 254, [10] := -256, [50] := 128, [51] := 9, [52] := 210, [54] := 1, [55] := 210, [60] := 25600, [61] := 9, [62] := 210, [64] := 17408, [66] := 210);
   N241 : DINT[1];
   N242 : DINT[2] := ([0] := -9, [1] := -9);
   N250 : DINT[100] := ([8] := 99, [10] := -256, [50] := -32640, [51] := 9, [52] := 200, [54] := 1, [55] := 200, [61] := 9, [62] := 200, [65] := 1, [66] := 200);
   N251 : DINT[100];
   N252 : DINT[100] := ([0] := -9, [1] := -9);
   N26 : DINT[33] := ([1] := 8, [10] := 38, [11] := 1, [30] := -15194, [31] := 8);
   N27 : DINT[50] := ([40] := 28176, [41] := 29344, [42] := 23976, [43] := 25960, [44] := 29304, [45] := 27664, [46] := 28928, [47] := 16);
   N28 : DINT[17] := ([0] := 124, [1] := 158, [2] := 937, [3] := 50, [4] := 9, [5] := 156, [6] := 3, [10] := 1000, [12] := 100);
   N7 : DINT[100] := ([0] := 5, [1] := 20, [2] := 20, [4] := 30000, [7] := 48, [8] := 48, [9] := 48, [10] := 53, [11] := 53, [12] := 43, [13] := 46, [14] := 46, [15] := 46, [16] := 51, [17] := 51, [18] := 46, [50] := 1, [51] := 1, [52] := 1, [53] := 1, [54] := 1, [55] := 1, [56] := 1, [57] := 1, [58] := 1, [59] := 1, [60] := 1, [61] := 1, [62] := 1, [93] := 9, [99] := 9);
   N_RECVING_PIT_GATE_AUTO : ALIAS FOR Local:0:I.Data.2;
   N_RECVING_PIT_GATE_CLOSE : ALIAS FOR Local:5:O.Data.5;
   N_RECVING_PIT_GATE_OPEN : ALIAS FOR Local:5:O.Data.4;
   NU : DINT;
   O10 : ALIAS FOR R1S0_AENTR:10:O.Data;
   O10_000_Bit00 : ALIAS FOR O10.0;
   O10_000_Bit01 : ALIAS FOR O10.1;
   O10_000_Bit02 : ALIAS FOR O10.2;
   O10_000_Bit03 : ALIAS FOR O10.3;
   O10_000_Bit04 : ALIAS FOR O10.4;
   O10_000_Bit05 : ALIAS FOR O10.5;
   O10_000_Bit06 : ALIAS FOR O10.6;
   O10_000_Bit07 : ALIAS FOR O10.7;
   O10_000_Bit08 : ALIAS FOR O10.8;
   O10_000_Bit09 : ALIAS FOR O10.9;
   O10_000_Bit10 : ALIAS FOR O10.10;
   O10_000_Bit11 : ALIAS FOR O10.11;
   O10_000_Bit12 : ALIAS FOR O10.12;
   O10_000_Bit13 : ALIAS FOR O10.13;
   O10_000_Bit14 : ALIAS FOR O10.14;
   O10_000_Bit15 : ALIAS FOR O10.15;
   O11 : ALIAS FOR R1S0_AENTR:11:O.Data;
   O11_000_Bit00 : ALIAS FOR O11.0;
   O11_000_Bit01 : ALIAS FOR O11.1;
   O11_000_Bit02 : ALIAS FOR O11.2;
   O11_000_Bit03 : ALIAS FOR O11.3;
   O11_000_Bit04 : ALIAS FOR O11.4;
   O11_000_Bit05 : ALIAS FOR O11.5;
   O11_000_Bit06 : ALIAS FOR O11.6;
   O11_000_Bit07 : ALIAS FOR O11.7;
   O11_000_Bit08 : ALIAS FOR O11.8;
   O11_000_Bit09 : ALIAS FOR O11.9;
   O11_000_Bit10 : ALIAS FOR O11.10;
   O11_000_Bit11 : ALIAS FOR O11.11;
   O11_000_Bit12 : ALIAS FOR O11.12;
   O11_000_Bit13 : ALIAS FOR O11.13;
   O11_000_Bit14 : ALIAS FOR O11.14;
   O12 : ALIAS FOR R1S0_AENTR:12:O.Data;
   O12_000_Bit00 : ALIAS FOR O12.0;
   O12_000_Bit01 : ALIAS FOR O12.1;
   O12_000_Bit02 : ALIAS FOR O12.2;
   O12_000_Bit03 : ALIAS FOR O12.3;
   O12_000_Bit04 : ALIAS FOR O12.4;
   O12_000_Bit05 : ALIAS FOR O12.5;
   O12_000_Bit06 : ALIAS FOR O12.6;
   O12_000_Bit08 : ALIAS FOR O12.8;
   O12_000_Bit09 : ALIAS FOR O12.9;
   O12_000_Bit10 : ALIAS FOR O12.10;
   O12_000_Bit11 : ALIAS FOR O12.11;
   O12_000_Bit12 : ALIAS FOR O12.12;
   O12_000_Bit13 : ALIAS FOR O12.13;
   O12_000_Bit14 : ALIAS FOR O12.14;
   O12_000_Bit15 : ALIAS FOR O12.15;
   O13 : ALIAS FOR R2S0_AENTR:1:O.Data;
   O13_000_Bit00 : ALIAS FOR O13.0;
   O13_000_Bit01 : ALIAS FOR O13.1;
   O13_000_Bit02 : ALIAS FOR O13.2;
   O13_000_Bit03 : ALIAS FOR O13.3;
   O13_000_Bit04 : ALIAS FOR O13.4;
   O13_000_Bit05 : ALIAS FOR O13.5;
   O13_000_Bit06 : ALIAS FOR O13.6;
   O13_000_Bit07 : ALIAS FOR O13.7;
   O13_000_Bit08 : ALIAS FOR O13.8;
   O13_000_Bit09 : ALIAS FOR O13.9;
   O13_000_Bit10 : ALIAS FOR O13.10;
   O13_000_Bit15 : ALIAS FOR O13.15;
   O16 : INT[12] := ([0] := 2#0000_1000_0101_1010, [1] := 2#0000_1000_0101_1010, [2] := 2#0000_1000_0101_1010, [3] := 2#0000_1000_0101_1010, [4] := 2#0000_1000_0101_1010, [5] := 2#0000_1000_0101_1010, [6] := 2#0000_1000_0101_1010, [7] := 2#0000_1000_0101_1010);
   O17 : INT[12] := ([0] := 2#0000_1000_0101_1010, [1] := 2#0000_1000_0101_1010, [2] := 2#0000_1000_0101_1010, [3] := 2#0000_1000_0101_1010, [4] := 2#0000_1000_0101_1010, [5] := 2#0000_1000_0101_1010, [6] := 2#0000_1000_0101_1010, [7] := 2#0000_1000_0101_1010);
   O18 : INT[12] := ([0] := 2#0000_1000_0101_1010, [1] := 2#0000_1000_0101_1010, [2] := 2#0000_1000_0101_1010, [3] := 2#0000_1000_0101_1010, [4] := 2#0000_1000_0101_1010, [5] := 2#0000_1000_0101_1010, [6] := 2#0000_1010_1001_1101, [7] := 2#0000_1010_1001_1101);
   O24 : INT[32] := ([7] := 2#0000_0000_1000_0010);
   O24_001_Bit00 : ALIAS FOR O24[1].0;
   O24_001_Bit01 : ALIAS FOR O24[1].1;
   O24_001_Bit02 : ALIAS FOR O24[1].2;
   O24_001_Bit03 : ALIAS FOR O24[1].3;
   O24_001_Bit04 : ALIAS FOR O24[1].4;
   O24_005_Bit00 : ALIAS FOR O24[5].0;
   O24_005_Bit01 : ALIAS FOR O24[5].1;
   O24_005_Bit02 : ALIAS FOR O24[5].2;
   O24_005_Bit03 : ALIAS FOR O24[5].3;
   O24_005_Bit04 : ALIAS FOR O24[5].4;
   O24_005_Bit05 : ALIAS FOR O24[5].5;
   O24_005_Bit06 : ALIAS FOR O24[5].6;
   O24_005_Bit07 : ALIAS FOR O24[5].7;
   O24_005_Bit08 : ALIAS FOR O24[5].8;
   O24_005_Bit09 : ALIAS FOR O24[5].9;
   O24_005_Bit10 : ALIAS FOR O24[5].10;
   O24_005_Bit11 : ALIAS FOR O24[5].11;
   O24_005_Bit12 : ALIAS FOR O24[5].12;
   O24_005_Bit15 : ALIAS FOR O24[5].15;
   O24_007_Bit00 : ALIAS FOR O24[7].0;
   O24_007_Bit01 : ALIAS FOR O24[7].1;
   O24_007_Bit04 : ALIAS FOR O24[7].4;
   O24_007_Bit05 : ALIAS FOR O24[7].5;
   O24_007_Bit06 : ALIAS FOR O24[7].6;
   O24_007_Bit07 : ALIAS FOR O24[7].7;
   O24_007_Bit10 : ALIAS FOR O24[7].10;
   O24_007_Bit11 : ALIAS FOR O24[7].11;
   O24_007_Bit12 : ALIAS FOR O24[7].12;
   O24_007_Bit13 : ALIAS FOR O24[7].13;
   O24_007_Bit14 : ALIAS FOR O24[7].14;
   O24_007_Bit8 : DINT;
   O25 : INT[32] := ([8] := 2#0100_0001_1101_1110, [9] := 2#0011_0111_0100_0010, [10] := 2#1110_0000_0100_0000, [11] := 2#0000_0000_0000_1010);
   O25_008_Bit00 : ALIAS FOR O25[8].0;
   O25_008_Bit01 : ALIAS FOR O25[8].1;
   O25_008_Bit02 : ALIAS FOR O25[8].2;
   O25_008_Bit03 : ALIAS FOR O25[8].3;
   O25_008_Bit04 : ALIAS FOR O25[8].4;
   O25_008_Bit06 : ALIAS FOR O25[8].6;
   O25_008_Bit07 : ALIAS FOR O25[8].7;
   O25_008_Bit08 : ALIAS FOR O25[8].8;
   O25_008_Bit09 : ALIAS FOR O25[8].9;
   O25_008_Bit10 : ALIAS FOR O25[8].10;
   O25_008_Bit12 : ALIAS FOR O25[8].12;
   O25_008_Bit13 : ALIAS FOR O25[8].13;
   O25_008_Bit14 : ALIAS FOR O25[8].14;
   O25_008_Bit15 : ALIAS FOR O25[8].15;
   O25_009_Bit00 : ALIAS FOR O25[9].0;
   O25_009_Bit01 : ALIAS FOR O25[9].1;
   O25_009_Bit02 : ALIAS FOR O25[9].2;
   O25_009_Bit03 : ALIAS FOR O25[9].3;
   O25_009_Bit04 : ALIAS FOR O25[9].4;
   O25_009_Bit05 : ALIAS FOR O25[9].5;
   O25_009_Bit06 : ALIAS FOR O25[9].6;
   O25_009_Bit07 : ALIAS FOR O25[9].7;
   O25_009_Bit08 : ALIAS FOR O25[9].8;
   O25_009_Bit09 : ALIAS FOR O25[9].9;
   O25_009_Bit10 : ALIAS FOR O25[9].10;
   O25_009_Bit11 : ALIAS FOR O25[9].11;
   O25_009_Bit12 : ALIAS FOR O25[9].12;
   O25_009_Bit13 : ALIAS FOR O25[9].13;
   O25_009_Bit14 : ALIAS FOR O25[9].14;
   O25_009_Bit15 : ALIAS FOR O25[9].15;
   O25_010_Bit00 : ALIAS FOR O25[10].0;
   O25_010_Bit01 : ALIAS FOR O25[10].1;
   O25_010_Bit02 : ALIAS FOR O25[10].2;
   O25_010_Bit03 : ALIAS FOR O25[10].3;
   O25_010_Bit04 : ALIAS FOR O25[10].4;
   O25_010_Bit05 : ALIAS FOR O25[10].5;
   O25_010_Bit06 : ALIAS FOR O25[10].6;
   O25_010_Bit07 : ALIAS FOR O25[10].7;
   O25_010_Bit08 : ALIAS FOR O25[10].8;
   O25_010_Bit09 : ALIAS FOR O25[10].9;
   O25_010_Bit10 : ALIAS FOR O25[10].10;
   O25_010_Bit11 : ALIAS FOR O25[10].11;
   O25_010_Bit12 : ALIAS FOR O25[10].12;
   O25_010_Bit13 : ALIAS FOR O25[10].13;
   O25_010_Bit14 : ALIAS FOR O25[10].14;
   O25_010_Bit15 : ALIAS FOR O25[10].15;
   O25_011_Bit00 : ALIAS FOR O25[11].0;
   O25_011_Bit01 : ALIAS FOR O25[11].1;
   O25_011_Bit03 : ALIAS FOR O25[11].3;
   O25_011_Bit14 : ALIAS FOR O25[11].14;
   O25_011_Bit15 : ALIAS FOR O25[11].15;
   O25_012_Bit00 : ALIAS FOR O25[12].0;
   O25_012_Bit01 : ALIAS FOR O25[12].1;
   O25_012_Bit02 : ALIAS FOR O25[12].2;
   O25_012_Bit03 : ALIAS FOR O25[12].3;
   O25_012_Bit04 : ALIAS FOR O25[12].4;
   O25_012_Bit05 : ALIAS FOR O25[12].5;
   O25_012_Bit06 : ALIAS FOR O25[12].6;
   O25_012_Bit07 : ALIAS FOR O25[12].7;
   O25_012_Bit08 : ALIAS FOR O25[12].8;
   O25_012_Bit09 : ALIAS FOR O25[12].9;
   O25_012_Bit10 : ALIAS FOR O25[12].10;
   O25_012_Bit11 : ALIAS FOR O25[12].11;
   O25_012_Bit12 : ALIAS FOR O25[12].12;
   O25_012_Bit13 : ALIAS FOR O25[12].13;
   O25_012_Bit14 : ALIAS FOR O25[12].14;
   O9 : ALIAS FOR R1S0_AENTR:9:O.Data;
   O9_000_Bit00 : ALIAS FOR O9.0;
   O9_000_Bit01 : ALIAS FOR O9.1;
   O9_000_Bit02 : ALIAS FOR O9.2;
   O9_000_Bit03 : ALIAS FOR O9.3;
   O9_000_Bit04 : ALIAS FOR O9.4;
   O9_000_Bit05 : ALIAS FOR O9.5;
   O9_000_Bit06 : ALIAS FOR O9.6;
   O9_000_Bit07 : ALIAS FOR O9.7;
   O9_000_Bit08 : ALIAS FOR O9.8;
   O9_000_Bit09 : ALIAS FOR O9.9;
   O9_000_Bit10 : ALIAS FOR O9.10;
   O9_000_Bit11 : ALIAS FOR O9.11;
   O9_000_Bit12 : ALIAS FOR O9.12;
   O9_000_Bit13 : ALIAS FOR O9.13;
   O9_000_Bit14 : ALIAS FOR O9.14;
   O9_000_Bit15 : ALIAS FOR O9.15;
   OLIVER_BIN : ALIAS FOR I4.8;
   OLIVER_SEP : ALIAS FOR I25[3].11;
   output_Bit : BOOL;
   Output_Bit_2 : BOOL;
   P10_ALARM : ALIAS FOR T4[97];
   P10_ALARM1 : ALIAS FOR T4[99];
   P10_AUTO_S : ALIAS FOR B3[5].10;
   P10_FLOW_A : ALIAS FOR N13[82];
   P10_FLOW_P : ALIAS FOR I24[21].8;
   P10_FLOW_P1 : ALIAS FOR C5[39];
   P10_FLW_OZ : ALIAS FOR N13[80];
   P10_MB : ALIAS FOR B12[10].2;
   P10_NO_FLO : ALIAS FOR B12[10].3;
   P10_OZ : ALIAS FOR N13[81];
   P10_RUN_AU : ALIAS FOR O24[5].9;
   P10_RUN_AU1 : ALIAS FOR B3[4].10;
   P10_SEC_SE : ALIAS FOR B17[1].10;
   P10_SEL_SW : ALIAS FOR I24[4].9;
   P10_SET : ALIAS FOR B12[10].0;
   P10_SPEED : ALIAS FOR N13[84];
   P10_STOP : ALIAS FOR B12[10].1;
   P11_RUN_AU : ALIAS FOR O24[5].10;
   P11_SEL_SW : ALIAS FOR I24[4].10;
   P12_RUN_AU : ALIAS FOR O24[5].11;
   P12_SEL_SW : ALIAS FOR I24[4].11;
   P1_ALARM_N : ALIAS FOR T4[81];
   P1_ALARM_N1 : ALIAS FOR T4[82];
   P1_AUTO_SE : ALIAS FOR B3[5].1;
   P1_FLOW_AN : ALIAS FOR N13[2];
   P1_FLOW_PL : ALIAS FOR C5[30];
   P1_FLOW_PU : ALIAS FOR I24[21].0;
   P1_FLW_OZ : ALIAS FOR N13[0];
   P1_MB : ALIAS FOR B12[1].2;
   P1_NO_FLOW : ALIAS FOR B12[1].3;
   P1_OZ : ALIAS FOR N13[1];
   P1_RUN_AUT : ALIAS FOR O24[5].0;
   P1_RUN_AUT1 : ALIAS FOR B3[4].1;
   P1_SEC_SEL : ALIAS FOR B17[1].1;
   P1_SEL_SW : ALIAS FOR I24[4].0;
   P1_SET : ALIAS FOR B12[1].0;
   P1_SPEED_O : ALIAS FOR N13[4];
   P1_STOP : ALIAS FOR B12[1].1;
   P2_ALARM_N : ALIAS FOR T4[83];
   P2_ALARM_N1 : ALIAS FOR T4[84];
   P2_AUTO_SE : ALIAS FOR B3[5].2;
   P2_FLOW_AN : ALIAS FOR N13[12];
   P2_FLOW_PL : ALIAS FOR C5[32];
   P2_FLOW_PU : ALIAS FOR I24[21].1;
   P2_FLW_OZ : ALIAS FOR N13[10];
   P2_MB : ALIAS FOR B12[2].2;
   P2_NO_FLOW : ALIAS FOR B12[2].3;
   P2_OZ : ALIAS FOR N13[11];
   P2_RUN_AUT : ALIAS FOR O24[5].1;
   P2_RUN_AUT1 : ALIAS FOR B3[4].2;
   P2_SEC_SEL : ALIAS FOR B17[1].2;
   P2_SEL_SW : ALIAS FOR I24[4].1;
   P2_SET : ALIAS FOR B12[2].0;
   P2_SPEED_O : ALIAS FOR N13[14];
   P2_STOP : ALIAS FOR B12[2].1;
   P3_ALARM_N : ALIAS FOR T4[85];
   P3_ALARM_N1 : ALIAS FOR T4[86];
   P3_AUTO_SE : ALIAS FOR B3[5].3;
   P3_FLOW_AN : ALIAS FOR N13[22];
   P3_FLOW_PL : ALIAS FOR C5[33];
   P3_FLOW_PU : ALIAS FOR I24[21].2;
   P3_FLW_OZ : ALIAS FOR N13[20];
   P3_MB : ALIAS FOR B12[3].2;
   P3_NO_FLOW : ALIAS FOR B12[3].3;
   P3_OZ : ALIAS FOR N13[21];
   P3_RUN_AUT : ALIAS FOR O24[5].2;
   P3_RUN_AUT1 : ALIAS FOR B3[4].3;
   P3_SEC_SEL : ALIAS FOR B17[1].3;
   P3_SEL_SW : ALIAS FOR I24[4].2;
   P3_SET : ALIAS FOR B12[3].0;
   P3_SPEED_O : ALIAS FOR N13[24];
   P3_STOP : ALIAS FOR B12[3].1;
   P4_ALARM_N : ALIAS FOR T4[87];
   P4_ALARM_N1 : ALIAS FOR T4[88];
   P4_AUTO_SE : ALIAS FOR B3[5].4;
   P4_FLOW_AN : ALIAS FOR N13[32];
   P4_FLOW_PL : ALIAS FOR C5[34];
   P4_FLOW_PU : ALIAS FOR I24[21].3;
   P4_FLW_OZ : ALIAS FOR N13[30];
   P4_MB : ALIAS FOR B12[4].2;
   P4_NO_FLOW : ALIAS FOR B12[4].3;
   P4_OZ : ALIAS FOR N13[31];
   P4_RUN_AUT : ALIAS FOR O24[5].3;
   P4_RUN_AUT1 : ALIAS FOR B3[4].4;
   P4_SEC_SEL : ALIAS FOR B17[1].4;
   P4_SEL_SW : ALIAS FOR I24[4].3;
   P4_SET : ALIAS FOR B12[4].0;
   P4_SPEED_O : ALIAS FOR N13[34];
   P4_STOP : ALIAS FOR B12[4].1;
   P5_ALARM_N : ALIAS FOR T4[89];
   P5_ALARM_N1 : ALIAS FOR T4[90];
   P5_AUTO_SE : ALIAS FOR B3[5].5;
   P5_FLOW_AN : ALIAS FOR N13[42];
   P5_FLOW_PL : ALIAS FOR C5[35];
   P5_FLOW_PU : ALIAS FOR I24[21].4;
   P5_FLW_OZ : ALIAS FOR N13[40];
   P5_MB : ALIAS FOR B12[5].2;
   P5_NO_FLOW : ALIAS FOR B12[5].3;
   P5_OZ : ALIAS FOR N13[41];
   P5_RUN_AUT : ALIAS FOR O24[5].4;
   P5_RUN_AUT1 : ALIAS FOR B3[4].5;
   P5_SEC_SEL : ALIAS FOR B17[1].5;
   P5_SEL_SW : ALIAS FOR I24[4].4;
   P5_SET : ALIAS FOR B12[5].0;
   P5_SPEED_O : ALIAS FOR N13[44];
   P5_STOP : ALIAS FOR B12[5].1;
   P6_ALARM_N : ALIAS FOR T4[91];
   P6_ALARM_N1 : ALIAS FOR T4[92];
   P6_AUTO_SE : ALIAS FOR B3[5].6;
   P6_FLOW_AN : ALIAS FOR N13[52];
   P6_FLOW_PL : ALIAS FOR C5[36];
   P6_FLOW_PU : ALIAS FOR I24[21].5;
   P6_FLW_OZ : ALIAS FOR N13[50];
   P6_MB : ALIAS FOR B12[6].2;
   P6_NO_FLOW : ALIAS FOR B12[6].3;
   P6_OZ : ALIAS FOR N13[51];
   P6_RUN_AUT : ALIAS FOR O24[5].5;
   P6_RUN_AUT1 : ALIAS FOR B3[4].6;
   P6_SEC_SEL : ALIAS FOR B17[1].6;
   P6_SEL_SW : ALIAS FOR I24[4].5;
   P6_SET : ALIAS FOR B12[6].0;
   P6_SPEED_O : ALIAS FOR N13[54];
   P6_STOP : ALIAS FOR B12[6].1;
   P7_ALARM_N : ALIAS FOR T4[93];
   P7_ALARM_N1 : ALIAS FOR T4[94];
   P7_AUTO_SE : ALIAS FOR B3[5].7;
   P7_FLOW_AN : ALIAS FOR N13[62];
   P7_FLOW_PL : ALIAS FOR C5[37];
   P7_FLOW_PU : ALIAS FOR I24[21].6;
   P7_FLW_OZ : ALIAS FOR N13[60];
   P7_MB : ALIAS FOR B12[7].2;
   P7_NO_FLOW : ALIAS FOR B12[7].3;
   P7_OZ : ALIAS FOR N13[61];
   P7_RUN_AUT : ALIAS FOR O24[5].6;
   P7_RUN_AUT1 : ALIAS FOR B3[4].7;
   P7_SEC_SEL : ALIAS FOR B17[1].7;
   P7_SEL_SW : ALIAS FOR I24[4].6;
   P7_SET : ALIAS FOR B12[7].0;
   P7_SPEED_O : ALIAS FOR N13[64];
   P7_STOP : ALIAS FOR B12[7].1;
   P8_ALARM_N : ALIAS FOR T4[95];
   P8_ALARM_N1 : ALIAS FOR T4[96];
   P8_AUTO_SE : ALIAS FOR B3[5].8;
   P8_FLOW_AN : ALIAS FOR N13[72];
   P8_FLOW_PL : ALIAS FOR C5[38];
   P8_FLOW_PU : ALIAS FOR I24[21].7;
   P8_FLW_OZ : ALIAS FOR N13[70];
   P8_MB : ALIAS FOR B12[8].2;
   P8_NO_FLOW : ALIAS FOR B12[8].3;
   P8_OZ : ALIAS FOR N13[71];
   P8_RUN_AUT : ALIAS FOR O24[5].7;
   P8_RUN_AUT1 : ALIAS FOR B3[4].8;
   P8_SEC_SEL : ALIAS FOR B17[1].8;
   P8_SEL_SW : ALIAS FOR I24[4].7;
   P8_SET : ALIAS FOR B12[8].0;
   P8_SPEED_O : ALIAS FOR N13[74];
   P8_STOP : ALIAS FOR B12[8].1;
   P9_RUN_AUT : ALIAS FOR O24[5].8;
   P9_SEC_SEL : ALIAS FOR B17[1].9;
   P9_SEL_SW : ALIAS FOR I24[4].8;
   P_RESET_AU : ALIAS FOR B3[4].0;
   PMP_15_OFF_DLY : REAL := 5.0;
   PMP_15_OFF_DLY_SCALE : REAL := 5000.0;
   PMP_15_ON_DLY : REAL := 5.0;
   PMP_15_ON_DLY_SCALE : REAL := 5000.0;
   PMP_15_TMR : TIMER := (PRE := 5000);
   PMP_15_TMR_2 : TIMER := (PRE := 5000);
   ProcessAll : BOOL;
   PUMP_13_RUN : ALIAS FOR R3M1_AENTR:3:O.8;
   PUMP_14_RUN : ALIAS FOR R3M1_AENTR:3:O.9;
   PUMP_15_AUTO : BOOL;
   PUMP_15_RUN : ALIAS FOR R3M1_AENTR:3:O.14;
   PUMP_NO_FL : ALIAS FOR B12[11].0;
   R6 : CONTROL[1];
   Rack24_1_Mode : BOOL := 1;
   RemoteAndcoAnalogIn : DINT[40] := ([1] := 9993, [3] := 10270, [4] := 5041, [5] := 7694, [7] := 9661, [9] := 3611, [10] := 9885, [11] := 8109, [12] := 10717, [13] := 7657, [14] := 9078, [15] := 8853, [19] := 9087, [20] := 9586);
   RSSql_MSG_BTR : INT;
   RSSql_MSG_BTR_DN : ALIAS FOR RSSql_MSG_BTR.0;
   RSSql_MSG_BTR_ER : ALIAS FOR RSSql_MSG_BTR.1;
   RSSql_MSG_Control : MESSAGE;
        MessageParameters(ServiceCode := 16#004d, LocalElement := spTicketTableBay1Wt, ...)
   RSSql_MSG_Data : DINT := 138;
   RSSql_MSG_En : BOOL;
   RSVIEW_ALA : ALIAS FOR B3[0].11;
   S : INT[83] := ([0] := 16#0004, [1] := 16#00de, [2] := 16#9032, [3] := 16#a005, [4] := 16#455e, [5] := 16#4000, [9] := 16#0002, [10] := 16#0032, [11] := 16#ffff, [12] := 16#ffff, [17] := 16#0002, [20] := 16#0001, [21] := 16#0008, [22] := 16#0006, [23] := 16#0005, [27] := 16#ffff, [28] := 16#ffff, [33] := 16#0208, [35] := 16#0030, [54] := 16#0021, [57] := 16#01f5, [58] := 16#0002, [59] := 16#0006, [60] := 16#0227, [61] := 16#0001, [62] := 16#0004, [63] := 16#0801, [64] := 16#0005, [65] := 16#0010, [66] := 16#0200);
   S24 : ALIAS FOR S[24];
   SCP_AOI : SCP_Inv[8] := ([0].In := 28184.0, [0].InRawMin := 12336.0, [0].InRawMax := 28816.0, [0].InEUMax := 3200.0, [0].Out := 122.71826, [1].In := 29344.0, [1].InRawMin := 10744.0, [1].InRawMax := 30320.0, [1].InEUMax := 3200.0, [1].Out := 159.54224, [2].In := 23976.0, [2].InRawMin := 9280.0, [2].InRawMax := 30064.0, [2].InEUMax := 3200.0, [2].Out := 937.3364, [3].In := 25960.0, [3].InRawMin := 7368.0, [3].InRawMax := 26256.0, [3].InEUMax := 3200.0, [3].Out := 50.148193, [4].In := 29296.0, [4].InRawMin := 9080.0, [4].InRawMax := 29360.0, [4].InEUMax := 3200.0, [4].Out := 10.098633, [5].In := 27664.0, [5].InRawMin := 8256.0, [5].InRawMax := 28656.0, [5].InEUMax := 3200.0, [5].Out := 155.60791, [6].In := 28928.0, [6].InRawMin := 11696.0, [6].InRawMax := 28944.0, [6].InEUMax := 3200.0, [6].Out := 2.9685059);
   Screen_Cancel : DINT;
   SCREENER_DRAG_START : BOOL;
   SCREENER_DRAG_STOP : BOOL;
   SCREENER_LEG_START : BOOL;
   SCREENER_LEG_STOP : BOOL;
   SCREENINGS : ALIAS FOR I7.15;
   Select_Cal_Bins : BOOL;
   Select_Clean_Bins : BOOL := 1;
   Select_Treat_Bins : BOOL;
   sendData : BOOL;
   sendData1 : BOOL;
   sendData_ONS : DINT;
   spBinGateRates : DINT[50] := ([11] := 86, [12] := 95, [13] := 79, [14] := 94, [15] := 93, [16] := 31, [17] := 79, [21] := 95, [22] := 83, [23] := 97, [24] := 90, [25] := 103, [26] := 99);
   spCapGrossWt : BOOL;
   spCapTareWt : BOOL;
   spCreateTicket : BOOL;
   spShowCreateTicketPB : BOOL;
   spTicketBinActive : DINT;
   spTicketBinSet : DINT;
   spTicketProcessing : BOOL;
   spTicketProcessStr : BOOL;
   spTicketTableBay1GrsWt : DINT;
   spTicketTableBay1Wt : DINT;
   spVAR_BINARRAY : STRING[50] := ([11] := '803001-Azimut-Certified - Limagrain  - HRW Seed Wheat', [12] := '883004-Lenetah-Certified -   - Barley Seed', [15] := '843002-Expresso-Certified-Monsanto -DNS Seed Wheat', [16] := '843005-Glee -Certified-WSU -DNS Seed Wheat', [17] := '843006-Kelse-Certified-WSU -DNS Seed Wheat', [22] := '843001-Buck Pronto-Certified-Limagrain -DNS Seed Wheat', [23] := '843004-SY 605-Certified-Sygenta Clearfield-DNS Seed Wheat', [24] := '803004-Keldin -Certified-Monsanto -HRW Seed Wheat', [25] := '843001-Buck Pronto-Certified-Limagrain -DNS Seed Wheat', [26] := '843003-Solano-Certified - Monsanto  - DNS Seed Wheat');
   sqlIndex : DINT;
   sqlIndex1 : DINT;
   sqlNewStartWeight : BOOL;
   sqlNewTreatment : BOOL;
   sqlNewTreatments_ONS : DINT;
   sqlNewVariety : BOOL;
   sqlNewVariety_ONS : DINT;
   sqlStartWtRecvd : DINT := 1;
   sqlTreatID : DINT;
   sqlTreatmentsRevd : DINT;
   sqlTreatRate : DINT;
   sqlTrtSendDelayTMR : TIMER := (PRE := 1000);
   sqlVaritiesRevd : DINT;
   sqlVarityID : DINT;
   sqlVarityRate : DINT;
   sqlVarSendDelayTMR : TIMER := (PRE := 1000);
   strEmptyVar : STRING := 'Empty';
   SURGE_BIN_HI : ALIAS FOR Local:0:I.Data.0;
   SURGE_BIN_LO : ALIAS FOR Local:0:I.Data.1;
   SWW_Index : DINT := 100;
   SWW_Variety_DB : Varieties_DB[100] := ([0].Id := 821001, [0].Name := 'ArtDeco', [0].ClassId := 1, [0].ClassType := 'Foundation', [0].MarketClassId := 82, [0].MarketClassType := 'SWW', [0].FullDecription := '821001  ArtDeco  Foundation  SWW', [1].Id := 822001, [1].Name := 'ArtDeco', [1].ClassId := 2, [1].ClassType := 'Registered', [1].MarketClassId := 82, [1].MarketClassType := 'SWW', [1].FullDecription := '822001  ArtDeco  Registered  SWW', [2].Id := 823001, [2].Name := 'ArtDeco', [2].ClassId := 3, [2].ClassType := 'Certified', [2].MarketClassId := 82, [2].MarketClassType := 'SWW', [2].FullDecription := '823001  ArtDeco  Certified  SWW', [3].Id := 821002, [3].Name := 'Huffman', [3].ClassId := 1, [3].ClassType := 'Foundation', [3].MarketClassId := 82, [3].MarketClassType := 'SWW', [3].FullDecription := '821002  Huffman  Foundation  SWW', [4].Id := 822002, [4].Name := 'Huffman', [4].ClassId := 2, [4].ClassType := 'Registered', [4].MarketClassId := 82, [4].MarketClassType := 'SWW', [4].FullDecription := '822002  Huffman  Registered  SWW', [5].Id := 823002, [5].Name := 'Huffman', [5].ClassId := 3, [5].ClassType := 'Certified', [5].MarketClassId := 82, [5].MarketClassType := 'SWW', [5].FullDecription := '823002  Huffman  Certified  SWW', [6].Id := 821003, [6].Name := 'WB 1035 CL Spring', [6].ClassId := 1, [6].ClassType := 'Foundation', [6].MarketClassId := 82, [6].MarketClassType := 'SWW', [6].FullDecription := '821003  WB 1035 CL Spring Foundation  SWW', [7].Id := 822003, [7].Name := 'WB 1035 CL Spring', [7].ClassId := 2, [7].ClassType := 'Registered', [7].MarketClassId := 82, [7].MarketClassType := 'SWW', [7].FullDecription := '822003  WB 1035 CL Spring  Registered  SWW', [8].Id := 823003, [8].Name := 'WB 1035 CL Spring', [8].ClassId := 3, [8].ClassType := 'Certified',
        [8].MarketClassId := 82, [8].MarketClassType := 'SWW', [8].FullDecription := '823003  WB 1035 CL Spring  Certified SWW');
   SWW_VarietySize : DINT := 100;
   SYMBOL : ALIAS FOR B3[0].0;
   SYMBOL_ANA : ALIAS FOR N10[1];
   T11 : TIMER[100] := ([0].PRE := 500, [0].ACC := 500, [0].EN := 1, [0].DN := 1, [1].PRE := 500, [1].ACC := 125, [1].EN := 1, [1].TT := 1, [3].PRE := 600000, [4].PRE := 1000, [5].PRE := 5000, [6].PRE := 5000, [7].PRE := 600000, [10].PRE := 5000, [11].PRE := 5000, [12].PRE := 5000, [13].PRE := 5000, [14].PRE := 5000, [15].PRE := 25000, [16].PRE := 5000, [17].PRE := 5000, [18].PRE := 5000, [19].PRE := 20000, [19].ACC := 20000, [19].EN := 1, [19].DN := 1);
   T11_AIR_SV : ALIAS FOR O9.0;
   T11_AIRSG : ALIAS FOR I1.0;
   T11_AIRSG1 : ALIAS FOR T4[0];
   T11_AIRSG2 : ALIAS FOR T4[1];
   T11_ASCII : ALIAS FOR B17[11].1;
   T11_ASSII : ALIAS FOR A16[112];
   T11_ASSII1 : ALIAS FOR A16[115];
   T11_AUTO_A : ALIAS FOR T4[61];
   T11_AUTO_A1 : ALIAS FOR T4[61].PRE;
   T11_AUTO_A2 : ALIAS FOR T4[61].ACC;
   T11_AUTO_M : ALIAS FOR B3[11].1;
   T11_AUTO_S : ALIAS FOR B3[11].14;
   T11_BINDIC : ALIAS FOR I4.11;
   T11_CAL_CL : ALIAS FOR B15[51].3;
   T11_CAL_LA : ALIAS FOR B15[51].2;
   T11_CAL_OP : ALIAS FOR B15[51].4;
   T11_CAL_ST : ALIAS FOR B15[51].1;
   T11_CLOSE : ALIAS FOR O9.1;
   T11_CLOSE1 : ALIAS FOR B3[11].9;
   T11_CLOSE2 : ALIAS FOR B3[11].11;
   T11_CORREC : ALIAS FOR F8[2];
   T11_DLY_TR : ALIAS FOR T4[0].PRE;
   T11_DLY_TR1 : ALIAS FOR T4[0].ACC;
   T11_DLY_TR2 : ALIAS FOR T4[1].PRE;
   T11_DLY_TR3 : ALIAS FOR T4[1].ACC;
   T11_FAULT : ALIAS FOR B3[11].15;
   T11_GATE_C : ALIAS FOR C5[11];
   T11_GATE_C1 : ALIAS FOR C5[11].PRE;
   T11_GATE_C2 : ALIAS FOR C5[11].ACC;
   T11_HOLD_A : ALIAS FOR B3[11].3;
   T11_HOLD_M : ALIAS FOR B3[11].6;
   T11_K_FACT : ALIAS FOR F8[1];
   T11_LOW_BI : ALIAS FOR B15[11].2;
   T11_MTR_GT : ALIAS FOR I1.2;
   T11_NO_PAS : ALIAS FOR B17[11].2;
   T11_NULL_V : ALIAS FOR A16[118];
   T11_NULL_V1 : ALIAS FOR A16[119];
   T11_OP_DEF : ALIAS FOR A16[116];
   T11_OP_DEF1 : ALIAS FOR A16[117];
   T11_OP_NAM : ALIAS FOR A16[113];
   T11_OP_NAM1 : ALIAS FOR A16[114];
   T11_OPEN_A : ALIAS FOR B3[11].8;
   T11_OPEN_M : ALIAS FOR O9.2;
   T11_OPEN_M1 : ALIAS FOR B3[11].10;
   T11_RELEAS : ALIAS FOR B3[11].5;
   T11_RESET : ALIAS FOR B3[11].7;
   T11_SET_AU : ALIAS FOR B3[11].2;
   T11_SET_DE : ALIAS FOR B3[2].0;
   T11_SET_LO : ALIAS FOR B3[11].13;
   T11_SET_MA : ALIAS FOR B3[11].12;
   T11_SET_NA : ALIAS FOR A16[110];
   T11_SET_NA1 : ALIAS FOR A16[111];
   T11_SET_NA2 : ALIAS FOR B17[11].0;
   T11_STOP_A : ALIAS FOR B3[11].4;
   T11_TREAT : ALIAS FOR B3[11].0;
   T11_TRT_MO : ALIAS FOR T4[41];
   T11_TRT_MO1 : ALIAS FOR T4[41].PRE;
   T11_TRT_MO2 : ALIAS FOR T4[41].ACC;
   T12_AIR_GA : ALIAS FOR I1.3;
   T12_AIR_SV : ALIAS FOR O9.3;
   T12_ASCII : ALIAS FOR B17[12].1;
   T12_ASSII : ALIAS FOR A16[122];
   T12_ASSII1 : ALIAS FOR A16[125];
   T12_AUTO_A : ALIAS FOR T4[62];
   T12_AUTO_A1 : ALIAS FOR T4[62].PRE;
   T12_AUTO_A2 : ALIAS FOR T4[62].ACC;
   T12_AUTO_M : ALIAS FOR B3[12].1;
   T12_AUTO_S : ALIAS FOR B3[12].14;
   T12_BINDIC : ALIAS FOR I4.12;
   T12_CAL_CL : ALIAS FOR B15[52].3;
   T12_CAL_LA : ALIAS FOR B15[52].2;
   T12_CAL_OP : ALIAS FOR B15[52].4;
   T12_CAL_ST : ALIAS FOR B15[52].1;
   T12_CLOSE : ALIAS FOR O9.4;
   T12_CLOSE1 : ALIAS FOR B3[12].9;
   T12_CLOSE2 : ALIAS FOR B3[12].11;
   T12_CORREC : ALIAS FOR F8[4];
   T12_DLY_TR : ALIAS FOR T4[2];
   T12_DLY_TR1 : ALIAS FOR T4[2].PRE;
   T12_DLY_TR2 : ALIAS FOR T4[2].ACC;
   T12_DLY_TR3 : ALIAS FOR T4[3];
   T12_DLY_TR4 : ALIAS FOR T4[3].PRE;
   T12_DLY_TR5 : ALIAS FOR T4[3].ACC;
   T12_FAULT : ALIAS FOR B3[12].15;
   T12_GATE_C : ALIAS FOR C5[12];
   T12_GATE_C1 : ALIAS FOR C5[12].PRE;
   T12_GATE_C2 : ALIAS FOR C5[12].ACC;
   T12_HOLD_A : ALIAS FOR B3[12].3;
   T12_HOLD_M : ALIAS FOR B3[12].6;
   T12_K_FACT : ALIAS FOR F8[3];
   T12_LOW_BI : ALIAS FOR B15[12].2;
   T12_METER : ALIAS FOR I1.5;
   T12_NO_PAS : ALIAS FOR B17[12].2;
   T12_NULL_V : ALIAS FOR A16[128];
   T12_NULL_V1 : ALIAS FOR A16[129];
   T12_OP_DEF : ALIAS FOR A16[126];
   T12_OP_DEF1 : ALIAS FOR A16[127];
   T12_OP_NAM : ALIAS FOR A16[123];
   T12_OP_NAM1 : ALIAS FOR A16[124];
   T12_OPEN_A : ALIAS FOR B3[12].8;
   T12_OPEN_M : ALIAS FOR O9.5;
   T12_OPEN_M1 : ALIAS FOR B3[12].10;
   T12_RELEAS : ALIAS FOR B3[12].5;
   T12_RESET : ALIAS FOR B3[12].7;
   T12_SET_AU : ALIAS FOR B3[12].2;
   T12_SET_DE : ALIAS FOR B3[2].1;
   T12_SET_LO : ALIAS FOR B3[12].13;
   T12_SET_MA : ALIAS FOR B3[12].12;
   T12_SET_NA : ALIAS FOR A16[120];
   T12_SET_NA1 : ALIAS FOR A16[121];
   T12_SET_NA2 : ALIAS FOR B17[12].0;
   T12_STOP_A : ALIAS FOR B3[12].4;
   T12_TREAT : ALIAS FOR B3[12].0;
   T12_TRT_MO : ALIAS FOR T4[42];
   T12_TRT_MO1 : ALIAS FOR T4[42].PRE;
   T12_TRT_MO2 : ALIAS FOR T4[42].ACC;
   T13_AIR_GA : ALIAS FOR I1.6;
   T13_AIR_SV : ALIAS FOR O9.6;
   T13_ASCII : ALIAS FOR B17[13].1;
   T13_ASSII : ALIAS FOR A16[132];
   T13_ASSII1 : ALIAS FOR A16[135];
   T13_AUTO_A : ALIAS FOR T4[63];
   T13_AUTO_A1 : ALIAS FOR T4[63].PRE;
   T13_AUTO_A2 : ALIAS FOR T4[63].ACC;
   T13_AUTO_M : ALIAS FOR B3[13].1;
   T13_AUTO_S : ALIAS FOR B3[13].14;
   T13_BINDIC : ALIAS FOR I4.13;
   T13_CAL_CL : ALIAS FOR B15[53].3;
   T13_CAL_LA : ALIAS FOR B15[53].2;
   T13_CAL_OP : ALIAS FOR B15[53].4;
   T13_CAL_ST : ALIAS FOR B15[53].1;
   T13_CLOSE : ALIAS FOR O9.7;
   T13_CLOSE1 : ALIAS FOR B3[13].9;
   T13_CLOSE2 : ALIAS FOR B3[13].11;
   T13_CORREC : ALIAS FOR F8[6];
   T13_DLY_TR : ALIAS FOR T4[4];
   T13_DLY_TR1 : ALIAS FOR T4[4].PRE;
   T13_DLY_TR2 : ALIAS FOR T4[4].ACC;
   T13_DLY_TR3 : ALIAS FOR T4[5];
   T13_DLY_TR4 : ALIAS FOR T4[5].PRE;
   T13_DLY_TR5 : ALIAS FOR T4[5].ACC;
   T13_FAULT : ALIAS FOR B3[13].15;
   T13_GATE_C : ALIAS FOR C5[13];
   T13_GATE_C1 : ALIAS FOR C5[13].PRE;
   T13_GATE_C2 : ALIAS FOR C5[13].ACC;
   T13_HOLD_A : ALIAS FOR B3[13].3;
   T13_HOLD_M : ALIAS FOR B3[13].6;
   T13_K_FACT : ALIAS FOR F8[5];
   T13_LOW_BI : ALIAS FOR B15[13].2;
   T13_MTR_GA : ALIAS FOR I1.8;
   T13_NO_PAS : ALIAS FOR B17[13].2;
   T13_NULL_V : ALIAS FOR A16[138];
   T13_NULL_V1 : ALIAS FOR A16[139];
   T13_OP_DEF : ALIAS FOR A16[136];
   T13_OP_DEF1 : ALIAS FOR A16[137];
   T13_OP_NAM : ALIAS FOR A16[133];
   T13_OP_NAM1 : ALIAS FOR A16[134];
   T13_OPEN_A : ALIAS FOR B3[13].8;
   T13_OPEN_M : ALIAS FOR O9.8;
   T13_OPEN_M1 : ALIAS FOR B3[13].10;
   T13_RELEAS : ALIAS FOR B3[13].5;
   T13_RESET : ALIAS FOR B3[13].7;
   T13_SET_AU : ALIAS FOR B3[13].2;
   T13_SET_DE : ALIAS FOR B3[2].2;
   T13_SET_LO : ALIAS FOR B3[13].13;
   T13_SET_MA : ALIAS FOR B3[13].12;
   T13_SET_NA : ALIAS FOR A16[130];
   T13_SET_NA1 : ALIAS FOR A16[131];
   T13_SET_NA2 : ALIAS FOR B17[13].0;
   T13_STOP_A : ALIAS FOR B3[13].4;
   T13_TREAT : ALIAS FOR B3[13].0;
   T13_TRT_MO : ALIAS FOR T4[43];
   T13_TRT_MO1 : ALIAS FOR T4[43].PRE;
   T13_TRT_MO2 : ALIAS FOR T4[43].ACC;
   T13C_AIR_G : ALIAS FOR O12.10;
   T13C_CLOSE : ALIAS FOR T22[6];
   T13C_CLOSE1 : ALIAS FOR T22[6].PRE;
   T13C_CLOSE2 : ALIAS FOR T22[6].ACC;
   T13C_GATE : ALIAS FOR B21[0].0;
   T13C_GATE1 : ALIAS FOR B21[0].1;
   T13C_GATE2 : ALIAS FOR B21[0].3;
   T13C_GATE3 : ALIAS FOR B21[0].4;
   T13C_GATE4 : ALIAS FOR B21[0].5;
   T13C_GATE5 : ALIAS FOR B21[0].6;
   T13C_GATE6 : ALIAS FOR B21[0].7;
   T13C_GATE7 : ALIAS FOR B21[0].8;
   T13C_GATE8 : ALIAS FOR B21[0].9;
   T13C_GATEC : ALIAS FOR B21[0].2;
   T13C_GATET : ALIAS FOR C5[2];
   T13C_SET_D : ALIAS FOR B21[70].14;
   T13C_TMR_A : ALIAS FOR C5[2].ACC;
   T13C_TMR_P : ALIAS FOR C5[2].PRE;
   T13C_TREAT : ALIAS FOR B21[70].10;
   T13C_TRT_M : ALIAS FOR T22[7];
   T13C_TRT_M1 : ALIAS FOR T22[7].PRE;
   T13C_TRT_M2 : ALIAS FOR T22[7].ACC;
   T13C_TRT_O : ALIAS FOR T22[5];
   T13C_TRT_O1 : ALIAS FOR T22[5].PRE;
   T13C_TRT_O2 : ALIAS FOR T22[5].ACC;
   T14_AIR_GT : ALIAS FOR I1.9;
   T14_AIR_SV : ALIAS FOR O9.9;
   T14_ASCII : ALIAS FOR B17[14].1;
   T14_ASSII : ALIAS FOR A16[142];
   T14_ASSII1 : ALIAS FOR A16[145];
   T14_AUTO_A : ALIAS FOR T4[64];
   T14_AUTO_A1 : ALIAS FOR T4[64].PRE;
   T14_AUTO_A2 : ALIAS FOR T4[64].ACC;
   T14_AUTO_M : ALIAS FOR B3[14].1;
   T14_AUTO_S : ALIAS FOR B3[14].14;
   T14_BINDIC : ALIAS FOR I4.14;
   T14_CAL_CL : ALIAS FOR B15[54].3;
   T14_CAL_LA : ALIAS FOR B15[54].2;
   T14_CAL_OP : ALIAS FOR B15[54].4;
   T14_CAL_ST : ALIAS FOR B15[54].1;
   T14_CLOSE : ALIAS FOR O9.10;
   T14_CLOSE1 : ALIAS FOR B3[14].9;
   T14_CLOSE2 : ALIAS FOR B3[14].11;
   T14_CORREC : ALIAS FOR F8[8];
   T14_DLY_TR : ALIAS FOR T4[6];
   T14_DLY_TR1 : ALIAS FOR T4[6].PRE;
   T14_DLY_TR2 : ALIAS FOR T4[6].ACC;
   T14_DLY_TR3 : ALIAS FOR T4[7];
   T14_DLY_TR4 : ALIAS FOR T4[7].PRE;
   T14_DLY_TR5 : ALIAS FOR T4[7].ACC;
   T14_FAULT : ALIAS FOR B3[14].15;
   T14_GATE_C : ALIAS FOR C5[14];
   T14_GATE_C1 : ALIAS FOR C5[14].PRE;
   T14_GATE_C2 : ALIAS FOR C5[14].ACC;
   T14_HOLD_A : ALIAS FOR B3[14].3;
   T14_HOLD_M : ALIAS FOR B3[14].6;
   T14_K_FACT : ALIAS FOR F8[7];
   T14_LOW_BI : ALIAS FOR B15[14].2;
   T14_MTR_GT : ALIAS FOR I1.11;
   T14_NO_PAS : ALIAS FOR B17[14].2;
   T14_NULL_V : ALIAS FOR A16[148];
   T14_NULL_V1 : ALIAS FOR A16[149];
   T14_OP_DEF : ALIAS FOR A16[146];
   T14_OP_DEF1 : ALIAS FOR A16[147];
   T14_OP_NAM : ALIAS FOR A16[143];
   T14_OP_NAM1 : ALIAS FOR A16[144];
   T14_OPEN_A : ALIAS FOR B3[14].8;
   T14_OPEN_M : ALIAS FOR O9.11;
   T14_OPEN_M1 : ALIAS FOR B3[14].10;
   T14_RELEAS : ALIAS FOR B3[14].5;
   T14_RESET : ALIAS FOR B3[14].7;
   T14_SET_AU : ALIAS FOR B3[14].2;
   T14_SET_DE : ALIAS FOR B3[2].3;
   T14_SET_LO : ALIAS FOR B3[14].13;
   T14_SET_MA : ALIAS FOR B3[14].12;
   T14_SET_NA : ALIAS FOR A16[140];
   T14_SET_NA1 : ALIAS FOR A16[141];
   T14_SET_NA2 : ALIAS FOR B17[14].0;
   T14_STOP_A : ALIAS FOR B3[14].4;
   T14_TREAT : ALIAS FOR B3[14].0;
   T14_TRT_MO : ALIAS FOR T4[44];
   T14_TRT_MO1 : ALIAS FOR T4[44].PRE;
   T14_TRT_MO2 : ALIAS FOR T4[44].ACC;
   T15_AIR_GT : ALIAS FOR I1.12;
   T15_AIR_SV : ALIAS FOR O9.12;
   T15_ASCII : ALIAS FOR B17[15].1;
   T15_ASSII : ALIAS FOR A16[152];
   T15_ASSII1 : ALIAS FOR A16[155];
   T15_AUTO_A : ALIAS FOR T4[65];
   T15_AUTO_A1 : ALIAS FOR T4[65].PRE;
   T15_AUTO_A2 : ALIAS FOR T4[65].ACC;
   T15_AUTO_M : ALIAS FOR B3[15].1;
   T15_AUTO_S : ALIAS FOR B3[15].14;
   T15_BINDIC : ALIAS FOR I4.15;
   T15_CAL_CL : ALIAS FOR B15[55].3;
   T15_CAL_LA : ALIAS FOR B15[55].2;
   T15_CAL_OP : ALIAS FOR B15[55].4;
   T15_CAL_ST : ALIAS FOR B15[55].1;
   T15_CLOSE : ALIAS FOR O9.13;
   T15_CLOSE1 : ALIAS FOR B3[15].9;
   T15_CLOSE2 : ALIAS FOR B3[15].11;
   T15_CORREC : ALIAS FOR F8[10];
   T15_FAULT : ALIAS FOR B3[15].15;
   T15_GATE_C : ALIAS FOR C5[15];
   T15_GATE_C1 : ALIAS FOR C5[15].PRE;
   T15_GATE_C2 : ALIAS FOR C5[15].ACC;
   T15_HOLD_A : ALIAS FOR B3[15].3;
   T15_HOLD_M : ALIAS FOR B3[15].6;
   T15_K_FACT : ALIAS FOR F8[9];
   T15_LOW_BI : ALIAS FOR B15[15].2;
   T15_MTR_GT : ALIAS FOR I1.14;
   T15_NO_PAS : ALIAS FOR B17[15].2;
   T15_NULL_V : ALIAS FOR A16[158];
   T15_NULL_V1 : ALIAS FOR A16[159];
   T15_OP_DEF : ALIAS FOR A16[156];
   T15_OP_DEF1 : ALIAS FOR A16[157];
   T15_OP_NAM : ALIAS FOR A16[153];
   T15_OP_NAM1 : ALIAS FOR A16[154];
   T15_OPEN_A : ALIAS FOR B3[15].8;
   T15_OPEN_M : ALIAS FOR O9.14;
   T15_OPEN_M1 : ALIAS FOR B3[15].10;
   T15_RELEAS : ALIAS FOR B3[15].5;
   T15_RESET : ALIAS FOR B3[15].7;
   T15_SET_AU : ALIAS FOR B3[15].2;
   T15_SET_DE : ALIAS FOR B3[2].4;
   T15_SET_LO : ALIAS FOR B3[15].13;
   T15_SET_MA : ALIAS FOR B3[15].12;
   T15_SET_NA : ALIAS FOR A16[150];
   T15_SET_NA1 : ALIAS FOR A16[151];
   T15_SET_NA2 : ALIAS FOR B17[15].0;
   T15_STOP_A : ALIAS FOR B3[15].4;
   T15_TREAT : ALIAS FOR B3[15].0;
   T15_TRT_MO : ALIAS FOR T4[45];
   T15_TRT_MO1 : ALIAS FOR T4[45].PRE;
   T15_TRT_MO2 : ALIAS FOR T4[45].ACC;
   T15_TRT_OF : ALIAS FOR T4[9];
   T15_TRT_OF1 : ALIAS FOR T4[9].PRE;
   T15_TRT_OF2 : ALIAS FOR T4[9].ACC;
   T15_TRT_ON : ALIAS FOR T4[8];
   T15_TRT_ON1 : ALIAS FOR T4[8].PRE;
   T15_TRT_ON2 : ALIAS FOR T4[8].ACC;
   T16_AIR_GA : ALIAS FOR I2.0;
   T16_AIR_SV : ALIAS FOR O10.0;
   T16_ASCII : ALIAS FOR B17[16].1;
   T16_ASSII : ALIAS FOR A16[162];
   T16_ASSII1 : ALIAS FOR A16[165];
   T16_AUTO_A : ALIAS FOR T4[66];
   T16_AUTO_A1 : ALIAS FOR T4[66].PRE;
   T16_AUTO_A2 : ALIAS FOR T4[66].ACC;
   T16_AUTO_M : ALIAS FOR B3[16].1;
   T16_AUTO_S : ALIAS FOR B3[16].14;
   T16_BINDIC : ALIAS FOR I4.9;
   T16_CAL_CL : ALIAS FOR B15[56].3;
   T16_CAL_LA : ALIAS FOR B15[56].2;
   T16_CAL_OP : ALIAS FOR B15[56].4;
   T16_CAL_ST : ALIAS FOR B15[56].1;
   T16_CLOSE : ALIAS FOR O10.1;
   T16_CLOSE1 : ALIAS FOR B3[16].9;
   T16_CLOSE2 : ALIAS FOR B3[16].11;
   T16_CORREC : ALIAS FOR F8[12];
   T16_FAULT : ALIAS FOR B3[16].15;
   T16_GATE_C : ALIAS FOR C5[16];
   T16_GATE_C1 : ALIAS FOR C5[16].PRE;
   T16_GATE_C2 : ALIAS FOR C5[16].ACC;
   T16_HOLD_A : ALIAS FOR B3[16].3;
   T16_HOLD_M : ALIAS FOR B3[16].6;
   T16_K_FACT : ALIAS FOR F8[11];
   T16_LOW_BI : ALIAS FOR B15[16].2;
   T16_METER : ALIAS FOR I2.2;
   T16_NO_PAS : ALIAS FOR B17[16].2;
   T16_NULL_V : ALIAS FOR A16[168];
   T16_NULL_V1 : ALIAS FOR A16[169];
   T16_OP_DEF : ALIAS FOR A16[166];
   T16_OP_DEF1 : ALIAS FOR A16[167];
   T16_OP_NAM : ALIAS FOR A16[163];
   T16_OP_NAM1 : ALIAS FOR A16[164];
   T16_OPEN_A : ALIAS FOR B3[16].8;
   T16_OPEN_M : ALIAS FOR O10.2;
   T16_OPEN_M1 : ALIAS FOR B3[16].10;
   T16_RELEAS : ALIAS FOR B3[16].5;
   T16_RESET : ALIAS FOR B3[16].7;
   T16_SET_AU : ALIAS FOR B3[16].2;
   T16_SET_DE : ALIAS FOR B3[2].5;
   T16_SET_LO : ALIAS FOR B3[16].13;
   T16_SET_MA : ALIAS FOR B3[16].12;
   T16_SET_NA : ALIAS FOR A16[160];
   T16_SET_NA1 : ALIAS FOR A16[161];
   T16_SET_NA2 : ALIAS FOR B17[16].0;
   T16_STOP_A : ALIAS FOR B3[16].4;
   T16_TREAT : ALIAS FOR B3[16].0;
   T16_TRT_MO : ALIAS FOR T4[46];
   T16_TRT_MO1 : ALIAS FOR T4[46].PRE;
   T16_TRT_MO2 : ALIAS FOR T4[46].ACC;
   T16_TRT_OF : ALIAS FOR T4[11];
   T16_TRT_OF1 : ALIAS FOR T4[11].PRE;
   T16_TRT_OF2 : ALIAS FOR T4[11].ACC;
   T16_TRT_ON : ALIAS FOR T4[10];
   T16_TRT_ON1 : ALIAS FOR T4[10].PRE;
   T16_TRT_ON2 : ALIAS FOR T4[10].ACC;
   T17_AIR_GA : ALIAS FOR I2.3;
   T17_AIR_SV : ALIAS FOR O10.3;
   T17_ASCII : ALIAS FOR B17[17].1;
   T17_ASSII : ALIAS FOR A16[172];
   T17_ASSII1 : ALIAS FOR A16[175];
   T17_AUTO_A : ALIAS FOR T4[67];
   T17_AUTO_A1 : ALIAS FOR T4[67].PRE;
   T17_AUTO_A2 : ALIAS FOR T4[67].ACC;
   T17_AUTO_M : ALIAS FOR B3[17].1;
   T17_AUTO_S : ALIAS FOR B3[17].14;
   T17_BINDIC : ALIAS FOR I4.10;
   T17_CAL_CL : ALIAS FOR B15[57].3;
   T17_CAL_LA : ALIAS FOR B15[57].2;
   T17_CAL_OP : ALIAS FOR B15[57].4;
   T17_CAL_ST : ALIAS FOR B15[57].1;
   T17_CLOSE : ALIAS FOR O10.4;
   T17_CLOSE1 : ALIAS FOR B3[17].9;
   T17_CLOSE2 : ALIAS FOR B3[17].11;
   T17_CORREC : ALIAS FOR F8[14];
   T17_FAULT : ALIAS FOR B3[17].15;
   T17_GATE_C : ALIAS FOR C5[17];
   T17_GATE_C1 : ALIAS FOR C5[17].PRE;
   T17_GATE_C2 : ALIAS FOR C5[17].ACC;
